(* IEC 61131-3 sources: daoli-st-library/DL_MathData, 454 files *)

(* ---- FC_DL_AccelUnitConvert.st ---- *)
(*==============================================================================
 * 组件名称 (Component)  : FC_DL_AccelUnitConvert
 * 所属子库 (Sublibrary) : DL_MathData ｜ 版本 (Version) : 1.0.0 ｜ 2026-11-23
 * 兼容性   (Platform)   : CODESYS 3.5+ / TwinCAT 3 / 汇川 InoProShop / 施耐德 Machine Expert
 *                         仅依赖 IEC 61131-3 算术运算符，零厂商私有库
 * 功能描述 (Function)   : 加速度单位互转（系数表驱动）：以 m/s² 为中介单位，
 *                         fHub = fValue × kSrc，fResult = fHub ÷ kDst；系数为编译期非零常量，
 *                         纯常量除法，结构性无除零。枚举源/目标越界一律由 CASE ... ELSE
 *                         拦截并返回 0 哨兵（禁静默换算）。
 *                         **重力常数口径**：标准重力加速度 g₀ = 9.80665 m/s²（ISO 80000-3 /
 *                         CGPM 1901 定义值），非本地纬度实测值；本件不做纬度修正。
 * 接口     (Interface)  : 输入 fValue 被换算加速度 [源单位]、eSrc 源单位、eDst 目标单位；
 *                         输出 fConverted 换算结果 [目标单位]、eErrCode（E_DL_AccConvErr）；
 *                         返回值 = 数值可信标志（TRUE = fConverted 可信）。
 * 边界     (Boundary)   : ① 加速度为矢量分量，负值合法（减速 / 反向），不设符号闸。
 *                         ② 单位枚举越域 → 故障级 eInvalidUnit，结果哨兵 0。
 *                         ③ 非有限双判（NaN / ±Inf），命中即故障级 eNonFinite。
 *                         ④ 中介值与结果各复检一次（四段式第四段）。
 *                         ⑤ 零值合法（自由落体失重即 0 g），置信息级 eZeroValue。
 *                         ⑥ 零全局耦合（无 GVL / VAR_EXTERNAL / 物理地址）。
 * 码表     (Codes)      : 本件不占用全局数字码位（R297 零码位范式）；出口为 BOOL + LREAL +
 *                         本文件内 enum E_DL_AccConvErr（全库唯一属主）。
 * 分工声明 (Scope)      : 速度归 FC_DL_SpeedUnitConvert，力归 FC_DL_ForceUnitConvert；
 *                         g 与 m/s² 属加速度量纲，本件专属。
 * 归属     (Ownership)  : E_DL_AccUnit / E_DL_AccConvErr 归属本文件（全库唯一属主，R264）。
 * 红线自检 (Redline)    : R1 ✓ 零 GVL ｜ R2 ✓ 零 %I/%Q ｜ R3 ✓ 纯 IEC ｜ R4 ✓ 非有限双判 +
 *                         CASE ELSE 枚举兜底 + 常量除法无除零 ｜ R5 ✓ 逐行同行双语注释
 *                         R6 ✓ CASE ELSE 兜底（无状态机相位） ｜ R7 N/A（无实例调用）
 * 修订历史 (Revision)   : 2026-11-23  v1.0.0  R78-B2 首版
 * 验收向量 (Acceptance) :
 *   A1 fValue=9.80665, eSrc=eMps2, eDst=eG → 1.0（容差 1E-12）；
 *   A2 fValue=1.0, eSrc=eG, eDst=eMps2 → 9.80665；
 *   A3 fValue=-2.0, eSrc=eMps2, eDst=eG → -0.20394324259558562（负值合法）；
 *   A4 fValue=5.0, eSrc=eMps2, eDst=非法值 7 → 0 哨兵, eInvalidUnit, 返回 FALSE；
 *   A5 fValue=0.0, eSrc=eG, eDst=eMps2 → 0.0, eZeroValue, 返回 TRUE。
 *============================================================================*)

(*-----------------------------------------------------------------------------
 * 枚举: E_DL_AccUnit（加速度单位表，归属本文件，全库唯一属主）
 *----------------------------------------------------------------------------*)
TYPE E_DL_AccUnit :
(
    eMps2 := 0,   // 米每二次方秒（中介单位） / Metre per second squared, hub unit
    eG    := 1    // 标准重力加速度（9.80665 m/s²） / Standard gravity, 9.80665 m/s²
);
END_TYPE

(*-----------------------------------------------------------------------------
 * 枚举: E_DL_AccConvErr（加速度换算出口码；信息级 = 0..9，故障级 = 10 起）
 *----------------------------------------------------------------------------*)
TYPE E_DL_AccConvErr :
(
    eOk          := 0,   // 信息级：换算完成 / Info: conversion completed
    eZeroValue   := 1,   // 信息级：零加速度（失重 / 静止） / Info: zero acceleration, result still trustworthy
    eInvalidUnit := 10,  // 故障级：单位枚举越域 / Fault: unit enum out of domain
    eNonFinite   := 11   // 故障级：输入或结果非有限 / Fault: non-finite input or result
);
END_TYPE

FUNCTION FC_DL_AccelUnitConvert : BOOL
VAR_INPUT
    fValue : LREAL;         // 被换算加速度 [源单位] / Acceleration value in the source unit
    eSrc   : E_DL_AccUnit;  // 源单位枚举 [-] / Source unit enum
    eDst   : E_DL_AccUnit;  // 目标单位枚举 [-] / Destination unit enum
END_VAR
VAR_OUTPUT
    fConverted : LREAL;           // 换算结果 [目标单位] / Converted result in the destination unit
    eErrCode   : E_DL_AccConvErr;  // 出口码 [-] / Outlet code
END_VAR
VAR
    _bBadValue : BOOL;   // 输入非有限标志 [-] / Non-finite input flag
    _fHub      : LREAL;  // 中介加速度值 [m/s²] / Hub acceleration value in metres per second squared
END_VAR
VAR CONSTANT
    DL_ACC_ZERO  : LREAL := 0.0;       // 零基准与零值判定基准 [-] / Zero base
    DL_ACC_MPS2  : LREAL := 1.0;       // m/s² → m/s² 恒等系数 [-] / Hub identity factor
    DL_ACC_G     : LREAL := 9.80665;   // g → m/s² 换算系数（标准重力） / Standard gravity factor
    DL_ACC_EPS   : LREAL := 1.0E-12;   // 零值判定容差 [-] / Zero-detection tolerance
END_VAR

(* —— 段 0：出口预置安全侧 —— *)
FC_DL_AccelUnitConvert := FALSE;                     // 返回值预置不可信 / Return preset not trustworthy
fConverted := DL_ACC_ZERO;                           // 结果哨兵 0 / Result sentinel
eErrCode   := E_DL_AccConvErr.eInvalidUnit;          // 预置最严码 / Preset strictest code

(* —— 段 1：非有限域闸（R79 双判） —— *)
_bBadValue := (fValue <> fValue) OR ((fValue - fValue) <> DL_ACC_ZERO);      // 输入非有限 / Input non-finite
IF _bBadValue THEN
    eErrCode := E_DL_AccConvErr.eNonFinite;          // 故障级码 / Fault-level code
    RETURN;
END_IF

(* —— 段 2：源单位 → 中介 m/s²（CASE ELSE 拦截越域，R6） —— *)
CASE eSrc OF
    E_DL_AccUnit.eMps2 :
        _fHub := fValue * DL_ACC_MPS2;               // 直通 / Hub pass-through
    E_DL_AccUnit.eG :
        _fHub := fValue * DL_ACC_G;                  // g × 9.80665 / Gravity scaled to metres per second squared
ELSE
    _fHub     := DL_ACC_ZERO;                        // 中介值回哨兵 / Hub back to sentinel
    eErrCode  := E_DL_AccConvErr.eInvalidUnit;       // 故障级：源单位越域 / Fault: source unit out of domain
    RETURN;
END_CASE

(* —— 段 3：中介 m/s² → 目标单位（除数为常量，均非零） —— *)
CASE eDst OF
    E_DL_AccUnit.eMps2 :
        fConverted := _fHub / DL_ACC_MPS2;           // ÷1 / Divide by identity
    E_DL_AccUnit.eG :
        fConverted := _fHub / DL_ACC_G;              // ÷9.80665 / Divide by standard gravity factor
ELSE
    fConverted := DL_ACC_ZERO;                       // 结果回哨兵 / Result back to sentinel
    eErrCode   := E_DL_AccConvErr.eInvalidUnit;      // 故障级：目标单位越域 / Fault: destination out of domain
    RETURN;
END_CASE

(* —— 段 4：中介值与结果复检（四段式第四段） —— *)
IF (_fHub <> _fHub) OR ((_fHub - _fHub) <> DL_ACC_ZERO)
    OR (fConverted <> fConverted) OR ((fConverted - fConverted) <> DL_ACC_ZERO) THEN
    fConverted := DL_ACC_ZERO;                       // 复检异常回哨兵 / Recheck failed: sentinel
    eErrCode   := E_DL_AccConvErr.eNonFinite;        // 故障级码 / Fault-level code
    RETURN;
END_IF

(* —— 段 5：成功出口（零值单列信息码） —— *)
IF (fValue < DL_ACC_EPS) AND (fValue > -DL_ACC_EPS) THEN
    eErrCode := E_DL_AccConvErr.eZeroValue;          // 信息级：零加速度 / Info: zero acceleration
ELSE
    eErrCode := E_DL_AccConvErr.eOk;                 // 信息级：换算完成 / Info: conversion completed
END_IF
FC_DL_AccelUnitConvert := TRUE;                      // 换算有效 / Conversion valid
END_FUNCTION

(* ---- FC_DL_AngleUnitConvert.st ---- *)
// ==============================================================================
// 组件名 Component  : FC_DL_AngleUnitConvert
// 分类   Category   : DL_MathData
// 前缀   Naming     : FC_DL_ ｜ b/f/e 类型前缀制（R265）
// 版本   Version    : 1.0.0
// 复杂度 Complexity  : 低
// 功能   Purpose    : 角度单位换算（度 / 弧度 / 梯度）：统一转 rad 中间量
//                      再转目标单位，任意两单位直换（deg → grad 系数
//                      200/180 经 rad 中转自动成立）。非有限输入拒绝
//                      （bValid = FALSE、fOut = 0.0）。
// 开源溯源 Origin    : 道莅原创（角度单位定义为公开计量常识，本实现
//                      clean-room，未复制任何源码行；与 TempUnitConvert /
//                      PressUnitConvert / FlowUnitConvert 同族单位换算
//                      组织口径）
// 许可证 License    : MIT
// 参考   Reference  : IEC 61131-3:2013 §6.6.2 CASE 语义；角度单位换算公开
//                      计量定义（借定义，不抄实现）
// 平台   Platform   : 纯 IEC 61131-3（CASE / LREAL 四则），三平台通用
// 依赖   Depends    : 无（零委托、零库件；换算系数常量预乘，运行期零除法）
// 分工声明 Split     : FC_DL_AngleDiffWrap（角差归一）与 FC_DL_WrapAngleDeg
//                      （角度回绕）与本件互引；本件只做单位换算（不改
//                      角度主值、不回绕），归一 / 回绕语义归各自属主（R216）。
// 归属 Ownership     : E_DL_AngUnit 属主为本文件（全库唯一定义，R264）；
//                      引用件只引用不重声明。
// ------------------------------------------------------------------
// 边界 Boundary     :
//   一 非有限闸：fVal 为 NaN（自反判 x <> x）或 ±Inf（差值自反判
//      (x - x) <> (x - x)）或幅值越 1e30 上界 → bValid = FALSE、
//      fOut = 0.0 早退（故障级 0749，R272 非有限防护）；
//   二 零除法面：四向系数全部预乘为常量（PI/180、180/PI、PI/200、
//      200/PI 编译期落定），运行期无除法（除零面结构性消除）；
//   三 枚举闸：eFrom / eTo 非法枚举值（CASE ELSE 兜底）→ bValid =
//      FALSE、fOut = 0.0 早退（与 0749 同形出口合并一码，R90 反证句：
//      现有输出组合不可区分两场景）；
//   四 纯函数：无记忆量、无定时器、无边沿实例，每调用重算；
//   五 无全局、无外部变量、无物理地址。
// 错误码 Codes      :
//   16#0001_0749【故障级】输入非有限或枚举非法（bValid = FALSE、
//                fOut = 0.0 早退）
//   注：本件引脚契约按任务定稿无独立 eErr 出口，故障语义经
//   bValid = FALSE + fOut = 0.0 组合表达。
// 验收 Acceptance   :
//   算法已证（脚本）：未跑 ｜ 编译器已证（三平台）：未跑
//   V1 180 deg → rad = 3.14159265358979；V2 1 rad → deg = 57.2957795
//   V3 200 grad → rad = 3.14159265358979；V4 180 deg → grad = 200（200/180 系数）
//   V5 fVal = NaN → bValid = FALSE、fOut = 0.0
//   V6 eFrom 非法枚举 → bValid = FALSE、fOut = 0.0
// 修订记录 Revision  :
//   2026-11-22  v1.0.0  R65 首版（批 2 · 序号 7）
// ==============================================================================
TYPE E_DL_AngUnit :
(
    eDeg  := 0, // 度 [deg]，一周 360 / degrees, 360 per turn
    eRad  := 1, // 弧度 [rad]，一周 2*PI / radians, two pi per turn
    eGrad := 2  // 梯度 [grad]，一周 400 / gradians, 400 per turn
);
END_TYPE

FUNCTION FC_DL_AngleUnitConvert : BOOL
VAR_INPUT
    fVal  : LREAL;               // 输入角值 [源单位] / the input angle in the source unit
    eFrom : E_DL_AngUnit;        // 源单位枚举 [单位] / the source unit
    eTo   : E_DL_AngUnit;        // 目标单位枚举 [单位] / the target unit
END_VAR
VAR_OUTPUT
    fOut   : LREAL;              // 输出角值 [目标单位]，无效时 0.0 / the output angle in the target unit, zero when invalid
    bValid : BOOL;               // 结果可用 [-]，非有限或枚举非法为 FALSE / the validity flag
END_VAR
VAR
    fRad : LREAL;                // 中间弧度量 [rad]（统一中转）/ the intermediate radian value
END_VAR
VAR CONSTANT
    DL_AUC_D2R  : LREAL := 0.0174532925199433;   // 度 → 弧度系数 [rad/deg]，PI/180 预乘 / the deg to rad factor, pi over one eighty
    DL_AUC_R2D  : LREAL := 57.2957795130823;     // 弧度 → 度系数 [deg/rad]，180/PI 预乘 / the rad to deg factor
    DL_AUC_G2R  : LREAL := 0.0157079632679490;   // 梯度 → 弧度系数 [rad/grad]，PI/200 预乘 / the grad to rad factor, pi over two hundred
    DL_AUC_R2G  : LREAL := 63.6619772367581;     // 弧度 → 梯度系数 [grad/rad]，200/PI 预乘 / the rad to grad factor
    DL_AUC_FMAX : LREAL := 1.0E30;               // 非有限筛查幅值上限 [源单位] / the finiteness screening cap
END_VAR

// 段 1｜返回值与全部出口预置（R45 四段式第一段）/ segment 1, the preset of the return and all outlets
FC_DL_AngleUnitConvert := FALSE; // 返回值预置假 / preset the return false
fOut   := 0.0;                   // 输出预置零 [目标单位] / preset the output zero
bValid := FALSE;                 // 有效标志预置假 / preset the validity false
fRad   := 0.0;                   // 中间量预置零 [rad] / preset the intermediate zero

// 段 2｜非有限闸（边界一：NaN 自反判 + Inf 差值自反判 + 幅值上界，R272）/ segment 2, the non finite gate
IF (fVal <> fVal) OR ((fVal - fVal) <> 0.0) OR (ABS(fVal) > DL_AUC_FMAX) THEN // 输入非有限 / the input non finite
    fOut   := 0.0;               // 输出归零 [目标单位] / zero the output
    bValid := FALSE;             // 故障级 0749：拒绝换算 / refuse the conversion
    RETURN;                      // 早退 / early return
END_IF

// 段 3｜源单位归一到 rad（边界三：CASE 带 ELSE 兜底）/ segment 3, the source unit normalization to radians
CASE eFrom OF
    E_DL_AngUnit.eDeg:           // 度 → rad / degrees to radians
        fRad := fVal * DL_AUC_D2R; // 乘 PI/180 系数 [rad] / multiply the deg to rad factor
    E_DL_AngUnit.eRad:           // 弧度直通 / radians pass through
        fRad := fVal;            // 中转量即输入 [rad] / the intermediate is the input
    E_DL_AngUnit.eGrad:          // 梯度 → rad / gradians to radians
        fRad := fVal * DL_AUC_G2R; // 乘 PI/200 系数 [rad] / multiply the grad to rad factor
    ELSE                         // 非法枚举拦截（边界三）/ an illegal enumeration
        fOut   := 0.0;           // 输出归零 / zero the output
        bValid := FALSE;         // 故障级 0749 同形出口（R90 合并）/ the merged fault outlet
        RETURN;                  // 早退 / early return
END_CASE

// 段 4｜rad 转目标单位（边界三：CASE 带 ELSE 兜底）/ segment 4, the radians to the target unit
CASE eTo OF
    E_DL_AngUnit.eDeg:           // rad → 度 / radians to degrees
        fOut := fRad * DL_AUC_R2D; // 乘 180/PI 系数 [deg] / multiply the rad to deg factor
    E_DL_AngUnit.eRad:           // rad 直通 / radians pass through
        fOut := fRad;            // 输出即中转量 [rad] / the output is the intermediate
    E_DL_AngUnit.eGrad:          // rad → 梯度 / radians to gradians
        fOut := fRad * DL_AUC_R2G; // 乘 200/PI 系数（deg → grad 经此链自动得 200/180）[grad] / the rad to grad factor
    ELSE                         // 非法枚举拦截（边界三）/ an illegal enumeration
        fOut   := 0.0;           // 输出归零 / zero the output
        bValid := FALSE;         // 故障级 0749 同形出口（R90 合并）/ the merged fault outlet
        RETURN;                  // 早退 / early return
END_CASE

// 段 5｜统一出口 / segment 5, the unified outlet
bValid := TRUE;                  // 结果可用 / the result usable
FC_DL_AngleUnitConvert := TRUE;  // 返回成功 / return success
END_FUNCTION

(* ---- FC_DL_AreaUnitConvert.st ---- *)
(*==============================================================================
 * 组件名称 (Component)  : FC_DL_AreaUnitConvert
 * 所属子库 (Sublibrary) : DL_MathData
 * 当前版本 (Version)    : 1.0.0
 * 兼容性   (Platform)   : CODESYS 3.5+ / TwinCAT 3 / 汇川 InoProShop / 施耐德 Machine Expert
 *                         仅依赖 IEC 61131-3 算术运算符，零厂商私有库
 * 功能描述 (Function)   : 面积单位换算（系数表驱动）：以平方米（m²）为中介单位，
 *                         fHub = fValue × kSrc，fResult = fHub ÷ kDst；系数为编译期
 *                         非零常量，纯常量除法，结构性无除零。
 *                         **量纲警告**：面积系数是长度系数的平方（mm² = 1E-6 m²、
 *                         ft² = 0.09290304 m²），不可与长度系数混用；本件显式使用
 *                         平方后的常量，禁止由长度族推导。
 *                         面积非负：负值判故障级 eNegativeValue 并回哨兵 0。
 * 接口     (Interface)  : 输入 fValue 被换算面积 [源单位]、eSrc 源单位、eDst 目标单位；
 *                         输出 fConverted 换算结果 [目标单位]、eErrCode（E_DL_AreaConvErr）；
 *                         返回值 = bValid 数值可信标志（TRUE = fConverted 可信）。
 * 边界     (Boundary)   : ① 属主边界：只做单位换算，不做体积 = 面积 × 行程 的推导。
 *                         ② 单位枚举越域 → 故障级 eInvalidUnit，结果哨兵 0。
 *                         ③ 非有限双判，命中即故障级 eNonFinite。
 *                         ④ 负面积 → 故障级 eNegativeValue（拒绝，不钳位）。
 *                         ⑤ 零值合法（info 级 eZeroValue）。结果与中介值各复检一次。
 *                         ⑥ 极小量纲提示：mm² 值域可极大（1 m² = 1E6 mm²），LREAL 尾数
 *                         53 位，最大可表 1.8E308，无溢出风险；但仍做非有限复检。
 *                         ⑦ 零全局耦合（无 GVL / VAR_EXTERNAL / 物理地址）。
 * 分工声明 (Scope)      : 与 `FC_DL_LengthUnitConvert` 分工：长度归那件，本件自带平方系数，
 *                         严禁调用长度件再平方（会引入两次舍入误差并破坏枚举域闸）。
 * 来源标签 (Source Tag) : 开源溯源：lgf-math 换算系数（公开物理常数，clean-room 重写）；许可证 MIT（仅参考语义，代码原创）
 * 码表     (Codes)      : 本件不占用全局数字码位；出口为 BOOL + LREAL +
 *                         本文件内定义 enum E_DL_AreaConvErr（全库唯一）。
 * 红线自检 (Redline)    : R1 ✓ 零 GVL/VAR_EXTERNAL ｜ R2 ✓ 零 %I/%Q/%M ｜ R3 ✓ 纯 IEC 61131-3
 *                         R4 ✓ 非有限双判 + 枚举域闸 + 常量除法无除零 + 负值拒绝 ｜ R5 ✓ 声明逐行同行双语注释
 *                         R6 N/A（纯函数无状态机） ｜ R7 N/A（无实例调用）
 * 修订历史 (Revision)   : 2026-11-23  v1.0.0  R77 首版（批次 B2 · 序号 14）
 * 验收向量 (Acceptance) : ① fValue=1.0, eSrc=eM2, eDst=eMm2 → 1×1.0 = 1 m2,
 *                         ÷1E-6 = 1000000.0 mm2（容差 1E-3）；
 *                         ② fValue=1.0, eSrc=eFt2, eDst=eM2 → 1×0.09290304 = 0.09290304 m2；
 *                         ③ fValue=1000000.0, eSrc=eMm2, eDst=eM2 → 1000000×1E-6 = 1.0 m2；
 *                         ④ fValue=-1.0, eSrc=eM2, eDst=eFt2 → 返回 FALSE, 0, eNegativeValue。
 *==============================================================================*)

(*-----------------------------------------------------------------------------
 * 枚举: E_DL_AreaUnit（面积单位表，归属 DL_MathData，与本件同文件，全库唯一属主）
 *----------------------------------------------------------------------------*)
TYPE E_DL_AreaUnit :
(
    eMm2 := 0,   // 平方毫米（1E-6 m2） / Square millimetre
    eM2  := 1,   // 平方米（中介单位） / Square metre, hub unit
    eFt2 := 2    // 平方英尺（0.09290304 m2，= 0.3048^2） / Square foot
);
END_TYPE

(*-----------------------------------------------------------------------------
 * 枚举: E_DL_AreaConvErr（面积换算错误码）
 *----------------------------------------------------------------------------*)
TYPE E_DL_AreaConvErr :
(
    eOk            := 0,   // 信息级：换算完成 / Info: conversion completed
    eZeroValue     := 1,   // 信息级：输入为零（合法） / Info: zero input, legal
    eInvalidUnit   := 2,   // 故障级：单位枚举越域 / Fault: unit enum out of domain
    eNonFinite     := 3,   // 故障级：输入非有限 / Fault: non-finite input
    eNegativeValue := 4    // 故障级：负面积 / Fault: negative area
);
END_TYPE

FUNCTION FC_DL_AreaUnitConvert : BOOL
VAR_INPUT
    fValue : LREAL;          // 被换算面积值 [源单位] / Area value in source unit
    eSrc   : E_DL_AreaUnit;  // 源单位枚举 [-] / Source unit enum
    eDst   : E_DL_AreaUnit;  // 目标单位枚举 [-] / Destination unit enum
END_VAR
VAR_OUTPUT
    fConverted : LREAL;            // 换算结果 [目标单位] / Converted result
    eErrCode   : E_DL_AreaConvErr; // 错误码出口 [-] / Error code outlet
END_VAR
VAR
    _bNonFin : BOOL;   // 输入非有限当拍标志 [-] / Non-finite input flag
    _fHub    : LREAL;  // 中介面积值 [m2] / Hub area value in square metres
END_VAR
VAR CONSTANT
    DL_AUC_MM2  : LREAL := 1.0E-6;      // mm2 → m2 换算系数（0.001^2） [m2/mm2] / square millimetre to square metre factor
    DL_AUC_M2   : LREAL := 1.0;         // m2 → m2 恒等系数 [m2/m2] / square metre identity factor
    DL_AUC_FT2  : LREAL := 0.09290304;  // ft2 → m2 换算系数（0.3048^2） [m2/ft2] / square foot to square metre factor
    DL_AUC_ZERO : LREAL := 0.0;         // 零值与非有限判零基准 [-] / Zero and non-finite base
END_VAR

(* —— 段 0：出口预置安全值 —— *)
FC_DL_AreaUnitConvert := FALSE;                    // 返回值预置无效 / Return preset invalid
fConverted := DL_AUC_ZERO;                         // 结果哨兵 0 / Result sentinel
eErrCode   := E_DL_AreaConvErr.eInvalidUnit;       // 预置最严码 / Preset strictest code

(* —— 段 1：非有限域闸（R79 双判） —— *)
_bNonFin := (fValue <> fValue) OR ((fValue - fValue) <> DL_AUC_ZERO);   // 非有限判定 / Non-finite test
IF _bNonFin THEN
    eErrCode := E_DL_AreaConvErr.eNonFinite;       // 故障级码 / Fault-level code
    RETURN;
END_IF

(* —— 段 2：负面积域闸 —— *)
IF fValue < DL_AUC_ZERO THEN
    eErrCode := E_DL_AreaConvErr.eNegativeValue;   // 故障级码 / Fault-level code
    RETURN;
END_IF

(* —— 段 3：源单位 → 中介平方米 —— *)
IF eSrc = E_DL_AreaUnit.eMm2 THEN
    _fHub := fValue * DL_AUC_MM2;                  // mm2 × 1E-6 / square millimetre scaled
ELSIF eSrc = E_DL_AreaUnit.eM2 THEN
    _fHub := fValue * DL_AUC_M2;                   // m2 直通 / square metre pass-through
ELSIF eSrc = E_DL_AreaUnit.eFt2 THEN
    _fHub := fValue * DL_AUC_FT2;                  // ft2 × 0.09290304 / square foot scaled
ELSE
    RETURN;                                        // 源单位越域 / Source unit out of domain
END_IF

(* —— 段 4：中介平方米 → 目标单位（常量除法，分母非零） —— *)
IF eDst = E_DL_AreaUnit.eMm2 THEN
    fConverted := _fHub / DL_AUC_MM2;              // ÷1E-6（放大 1e6，注意量纲） / Divide by square millimetre factor
ELSIF eDst = E_DL_AreaUnit.eM2 THEN
    fConverted := _fHub / DL_AUC_M2;               // ÷1 / Divide by identity
ELSIF eDst = E_DL_AreaUnit.eFt2 THEN
    fConverted := _fHub / DL_AUC_FT2;              // ÷0.09290304 / Divide by square foot factor
ELSE
    eErrCode   := E_DL_AreaConvErr.eInvalidUnit;   // 目标单位越域 / Destination out of domain
    fConverted := DL_AUC_ZERO;
    RETURN;
END_IF

(* —— 段 5：结果非有限复检兜底（量级放大 1e6 后必须复检） —— *)
IF (fConverted <> fConverted) OR ((fConverted - fConverted) <> DL_AUC_ZERO) THEN
    fConverted := DL_AUC_ZERO;                     // 复检异常回哨兵 / Recheck failed: sentinel
    eErrCode   := E_DL_AreaConvErr.eNonFinite;     // 故障级码 / Fault-level code
    RETURN;
END_IF

(* —— 段 6：成功出口 —— *)
IF fValue = DL_AUC_ZERO THEN
    eErrCode := E_DL_AreaConvErr.eZeroValue;       // 信息级：零值 / Info: zero value
ELSE
    eErrCode := E_DL_AreaConvErr.eOk;              // 信息级成功 / Info success
END_IF
FC_DL_AreaUnitConvert := TRUE;                     // 换算有效 / Conversion valid

END_FUNCTION

(* ---- FC_DL_CharCodeConvert.st ---- *)
(*
    FC_DL_CharCodeConvert —— 单字符 ↔ 字符码双向换算原子
    ------------------------------------------------------------------
    组件名称  : FC_DL_CharCodeConvert
    分类      : DL_MathData / CharCode
    前缀      : FC_DL_
    版本      : 1.0.0
    溯源      : IEC 61131-3 标准语义的道莅防御性实现（单字符与码值的
                双向映射原子，映射内核 = 定长字符表 + 标准 MID / FIND
                检索，零内建转换链依赖）；实现 / 引脚名 / 码位 100% 自有；
                clean-room 声明 —— 零代码行复制，无闭源参考。
    平台      : 纯 IEC 61131-3（Standard.library: LEN / MID / FIND），
                CODESYS 3.5 / TwinCAT 3 / InoProShop / Machine Expert 通用
    作者      : 道莅代码库 · PLC编程专家（R72 构建轮 · 批 2 · 序号 4）
    ------------------------------------------------------------------
    功能说明  : 单字符与字符码（0~255）双向换算。真实工况：HMI 键盘映射、
                协议字符组装、标签打印机字符转义。选向由 eMode 枚举显式
                给出，未选方向出口置确定值（空串 / 0），绝不残留旧值。
                判据链顺序：
                ① eCharToCode 向：串长域闸（LEN <> 1 → 拒收信息级，空串 /
                   多字符同样拒收）→ LO / HI 双表 FIND 检索（先 LO 后 HI，
                   命中即回码值）→ 双表全未命中 → 防御性拒收（结构性不可达，
                   表覆盖 1..255 全字节）；
                ② eCodeToChar 向：码域闸（uCodeIn > 255 → 故障级早退）→
                   码 0 = 串终结符，回执空串（忠实语义，声明口径）→ 码
                   1..127 查 LO 表（位置 = 码值）、码 128..255 查 HI 表
                   （位置 = 码值 − 127）；
                ③ 选向枚举漏项由 CASE ELSE 兜底（拒收信息级，双出口置
                   确定值）。
                扩展 ASCII 披露（128~255）：本件只保证**码值回执**的字节级
                正确性，不保证三平台对 $80~$FF 的渲染 / 显示一致（字体与
                代码页差异属显示层语义），头注释声明披露。
                交付门槛（R64 口径）：MID / FIND 对 $80~$FF 字节的检索行为
                须在 CODESYS / TwinCAT / InoProShop 三平台各编译验证一次。
    错误码    : 16#0002_3906 码域越界（uCodeIn > 255），双出口置确定值空串/0
                            —— 故障级
                16#0002_3907 串长域闸拒收（LEN <> 1，空串 / 多字符同拒）
                            —— 信息级，不置 bError（R45）
                16#0002_3908 选向枚举漏项（CASE ELSE 兜底拒收）—— 信息级，
                            不置 bError
                加码反证句（R90）：3906 由「故障级 + 双出口确定值」唯一观测；
                3907 与 3908 在输出组合上不可分（同为拒收），但成因互斥
                （串长 vs 选向）且调用方可自证入参，故按成因分立两码，
                拒绝合并导致选向错误被误报为串长错误。
    码位总账  : 16#0002_3906 用 ｜ 16#0002_3907 用 ｜ 16#0002_3908 用
    状态机    : 无顺序状态机；选向用 CASE + ELSE 兜底（非法枚举值拦截），
                枚举成员初值一律 :=（红线 4）
    边界与披露: 一 无定时器 / 无沿检测实例 / 无数组下标 / 无除法，周期安全
                   规则 N/A；
                二 零全局变量、零 VAR_EXTERNAL、零物理地址；
                三 域闸逐项点名（R272）：uCodeIn 码域闸覆盖 0~255 全段
                   （0 与 255 两端点各推一条向量）；sCharIn 串长闸覆盖
                   0 / 1 / 多字符三态；
                四 双出口默认值纪律：未选向 / 拒收路径 sCharOut = ''、
                   uCodeOut = 0 确定值，绝不残留旧值（R256）；
                五 字符表覆盖声明：LO 表覆盖码 1..127、HI 表覆盖码 128..255、
                   码 0 按串终结符语义回执空串——三段并起覆盖 0..255 全域，
                   无缺口；
                六 与 FC_DL_HexStringToBytes / FC_DL_DwordToHexString 分工
                   互引：那两件是文本 ↔ 字节块，本件是单字符 ↔ 码值原子，
                   不互代；
                七 依赖声明：仅 Standard.library（LEN / MID / FIND），
                   零厂商方言。
    验收向量  : V1 eCodeToChar，uCodeIn = 0 → 空串（终结符语义）；
                V2 eCodeToChar，uCodeIn = 65 → 'A'；V3 eCodeToChar，
                uCodeIn = 255 → '$FF' 字符；V4 eCodeToChar，uCodeIn = 256
                → 3906 故障级；V5 eCharToCode，'A' → 65；
                V6 eCharToCode，'' 或 'AB' → 3907 拒收；
                V7 eCharToCode，' '（空格，码 32）→ 32。
                算法已证（脚本）：未跑 ｜ 编译器已证（三平台）：未跑
    修订记录  : 2026-11-23 v1.0.0 首次入库（R72 构建轮 · 批 2 · 序号 4）
*)
TYPE E_DL_CharCodeMode :
(
    eCharToCode := 0,                      // 选向：字符 → 码值 / the direction char to code
    eCodeToChar := 1                       // 选向：码值 → 字符 / the direction code to char
);
END_TYPE

FUNCTION FC_DL_CharCodeConvert : BOOL
VAR_INPUT
    eMode    : E_DL_CharCodeMode;          (* 换算方向选向，[选向枚举] / the conversion direction selector *)
    sCharIn  : STRING;                     (* 字符输入（eCharToCode 向用），[串]，串长闸限 1 字符 / the char input, gated to one char *)
    uCodeIn  : UINT;                       (* 码值输入（eCodeToChar 向用），[码]，域 0~255 / the code input, domain 0 to 255 *)
END_VAR
VAR_OUTPUT
    sCharOut  : STRING(1);                 (* 字符出口（未选向 / 拒收时为空串确定值）[串] / the char outlet, empty when rejected *)
    uCodeOut  : UINT;                      (* 码值出口（未选向 / 拒收时为 0 确定值）[码] / the code outlet, zero when rejected *)
    bValid    : BOOL;                      (* 输出可用标志，拒收 / 故障为 FALSE / the outputs usable flag *)
    bError    : BOOL;                      (* 故障标志，仅故障级码置位（R45 配对）/ the fault flag *)
    nInfoCode : UDINT;                     (* 信息 / 错误码，0 = 正常 / the info or error id *)
END_VAR
VAR CONSTANT
    DL_CHC_TAB_LO : STRING(127) := '$01$02$03$04$05$06$07$08$09$0A$0B$0C$0D$0E$0F$10$11$12$13$14$15$16$17$18$19$1A$1B$1C$1D$1E$1F !"$24%&$27()*+,-./0123456789:;<=>?@ABCDEFGHIJKLMNOPQRSTUVWXYZ[\]^_`abcdefghijklmnopqrstuvwxyz{|}~$7F'; (* 码 1..127 字符表（位置 p = 码 p），$24 = '$'，$27 = ''' / the low char table, position p equals code p *)
    DL_CHC_TAB_HI : STRING(128) := '$80$81$82$83$84$85$86$87$88$89$8A$8B$8C$8D$8E$8F$90$91$92$93$94$95$96$97$98$99$9A$9B$9C$9D$9E$9F$A0$A1$A2$A3$A4$A5$A6$A7$A8$A9$AA$AB$AC$AD$AE$AF$B0$B1$B2$B3$B4$B5$B6$B7$B8$B9$BA$BB$BC$BD$BE$BF$C0$C1$C2$C3$C4$C5$C6$C7$C8$C9$CA$CB$CC$CD$CE$CF$D0$D1$D2$D3$D4$D5$D6$D7$D8$D9$DA$DB$DC$DD$DE$DF$E0$E1$E2$E3$E4$E5$E6$E7$E8$E9$EA$EB$EC$ED$EE$EF$F0$F1$F2$F3$F4$F5$F6$F7$F8$F9$FA$FB$FC$FD$FE$FF'; (* 码 128..255 字符表（位置 p = 码 127 + p），只保证码值回执不保证显示 / the high char table, position p equals code 127 plus p *)
    DL_CHC_ONE    : INT  := 1;             (* 检索步进与串长基准 [个] / the search step and the length base *)
    DL_CHC_SPLIT  : UINT := 127;           (* LO / HI 表码值分界 [码] / the code split between the tables *)
    DL_CHC_CMAX   : UINT := 255;           (* 码域上界 [码] / the code domain upper bound *)
    DL_CHC_ZERO   : UINT := 0;             (* 码零哨兵（终结符语义）[码] / the zero code sentinel *)
    DL_CHC_ZEROI  : INT  := 0;             (* 检索未命中哨兵 [位置] / the not found sentinel *)
END_VAR
VAR
    nLen  : INT;                           (* 输入串长 [个] / the input string length *)
    nPos  : INT;                           (* FIND 检索命中位置（LO 表）[位置] / the FIND hit position in the low table *)
    nPosH : INT;                           (* FIND 检索命中位置（HI 表）[位置] / the FIND hit position in the high table *)
END_VAR

// 段 1｜返回值与双出口预置（统一出口预置，R256）/ segment 1, preset the return and the dual outlets
FC_DL_CharCodeConvert := FALSE;          // 故障缺省返回不可用 / the fault default is unusable
sCharOut  := '';                         // 字符出口预置空串确定值 / preset the char outlet to the empty string
uCodeOut  := DL_CHC_ZERO;                // 码值出口预置零确定值 / preset the code outlet to zero
bValid    := FALSE;                      // 可用标志预清零 / preset the usable flag false
bError    := FALSE;                      // 故障标志预清零 / preset the fault flag false
nInfoCode := 0;                          // 码位预置无错 / preset the code to zero
nLen  := 0;                              // 串长中间量清零 / clear the length temporary
nPos  := DL_CHC_ZEROI;                   // 检索位置清零 / clear the hit position
nPosH := DL_CHC_ZEROI;                   // 检索位置清零 / clear the hit position

// 段 2｜选向分发（CASE + ELSE 兜底，非法枚举值拦截，红线 4）/ segment 2, the direction dispatch with the ELSE guard
CASE eMode OF

    E_DL_CharCodeMode.eCharToCode:       // 字符 → 码值向 / the char to code direction
        nLen := LEN(sCharIn);            // 串长闸取样 / sample the input length
        IF nLen <> DL_CHC_ONE THEN       // 空串或多字符一律拒收（串长域闸）/ empty or multi char rejected
            nInfoCode := 16#0002_3907;   // 信息级：串长闸拒收 / info level: the length gate rejection
            bError := FALSE;             // 信息级不置故障（R45）/ info level never raises a fault
            bValid := FALSE;             // 输出不可用 / the outputs unusable
            sCharOut := '';              // 双出口确定值（R256）/ the deterministic outlets
            uCodeOut := DL_CHC_ZERO;     // 双出口确定值 / the deterministic outlets
            RETURN;                      // 结构早退 / structural exit
        END_IF
        nPos := FIND(DL_CHC_TAB_LO, sCharIn); // LO 表检索（位置 p = 码 p）/ search the low table
        IF nPos > DL_CHC_ZEROI THEN      // LO 表命中 / a low table hit
            uCodeOut := INT_TO_UINT(nPos); // 码值 = 位置 / the code equals the position
        ELSE                             // LO 未命中转 HI 表 / fall through to the high table
            nPosH := FIND(DL_CHC_TAB_HI, sCharIn); // HI 表检索（位置 p = 码 127 + p）/ search the high table
            IF nPosH > DL_CHC_ZEROI THEN // HI 表命中 / a high table hit
                uCodeOut := INT_TO_UINT(nPosH + UINT_TO_INT(DL_CHC_SPLIT)); // 码值 = 位置 + 127 / the code equals position plus 127
            ELSE                         // 双表全未命中（表覆盖 1..255 全字节，结构性不可达防御收口）/ both tables missed, unreachable
                nInfoCode := 16#0002_3907; // 信息级：检索失败按拒收口径 / info level: the search failure rejection
                bValid := FALSE;         // 输出不可用 / unusable
                sCharOut := '';          // 双出口确定值 / the deterministic outlets
                uCodeOut := DL_CHC_ZERO; // 双出口确定值 / the deterministic outlets
                RETURN;                  // 结构早退 / exit
            END_IF
        END_IF
        bValid := TRUE;                  // 换算成功 / the conversion succeeded

    E_DL_CharCodeMode.eCodeToChar:       // 码值 → 字符向 / the code to char direction
        IF uCodeIn > DL_CHC_CMAX THEN    // 码域闸（>255 越域）/ the code domain gate
            nInfoCode := 16#0002_3906;   // 故障级：码域越界 / fault level: the code domain violation
            bError := TRUE;              // R45 配对置故障标志 / paired with the fault flag
            bValid := FALSE;             // 输出不可用 / unusable
            sCharOut := '';              // 双出口确定值 / the deterministic outlets
            uCodeOut := DL_CHC_ZERO;     // 双出口确定值 / the deterministic outlets
            RETURN;                      // 结构早退 / exit
        END_IF
        uCodeOut := uCodeIn;             // 码值回执（选向确认）/ echo the code
        IF uCodeIn = DL_CHC_ZERO THEN    // 码 0 = 串终结符，忠实回执空串 / code zero is the terminator, faithful empty
            sCharOut := '';              // 空串出口 / the empty outlet
        ELSIF uCodeIn <= DL_CHC_SPLIT THEN // 码 1..127 查 LO 表 / the low table range
            nPos := UINT_TO_INT(uCodeIn); // 位置 = 码值（LO 表 1 起）/ the position equals the code
            sCharOut := MID(DL_CHC_TAB_LO, nPos, DL_CHC_ONE); // 取单字符 / pick the single char
        ELSE                             // 码 128..255 查 HI 表 / the high table range
            nPos := UINT_TO_INT(uCodeIn) - UINT_TO_INT(DL_CHC_SPLIT); // 位置 = 码值 − 127 / the position equals code minus 127
            sCharOut := MID(DL_CHC_TAB_HI, nPos, DL_CHC_ONE); // 取单字符 / pick the single char
        END_IF
        bValid := TRUE;                  // 换算成功 / the conversion succeeded

    ELSE                                 // 选向枚举漏项兜底（红线 4）/ the unknown direction guard
        nInfoCode := 16#0002_3908;       // 信息级：选向未知拒收 / info level: the unknown direction rejection
        bError := FALSE;                 // 信息级不置故障（R45）/ info level never raises a fault
        bValid := FALSE;                 // 输出不可用 / unusable
        sCharOut := '';                  // 双出口确定值 / the deterministic outlets
        uCodeOut := DL_CHC_ZERO;         // 双出口确定值 / the deterministic outlets

END_CASE

// 段 3｜统一出口 / segment 3, the unified outlet
FC_DL_CharCodeConvert := bValid;         // 返回值与 bValid 同源（R191 名实双出口）/ the return shares its source with bValid
END_FUNCTION

(* ---- FC_DL_CircleFit3Pt.st ---- *)
(*==============================================================================
 * 组件名称 (Component)  : FC_DL_CircleFit3Pt
 * 所属子库 (Sublibrary) : DL_MathData
 * 当前版本 (Version)    : 1.0.0
 * 兼容性   (Platform)   : CODESYS 3.5+ / TwinCAT 3 / 汇川 InoProShop / 施耐德 Machine Expert
 *                         仅依赖 Standard.library（SQRT / ABS），零厂商私有库
 * 功能描述 (Function)   : 三点定圆（外接圆解析解，代数行列式法）：
 *                           D  = 2×[x1(y2−y3) + x2(y3−y1) + x3(y1−y2)]
 *                           Ux = [(x1²+y1²)(y2−y3) + (x2²+y2²)(y3−y1)
 *                                 + (x3²+y3²)(y1−y2)] ÷ D
 *                           Uy = [(x1²+y1²)(x3−x2) + (x2²+y2²)(x1−x3)
 *                                 + (x3²+y3²)(x2−x1)] ÷ D
 *                           R  = SQRT((x1−Ux)² + (y1−Uy)²)
 *                         |D| < 共线容差判三点共线（叉积绝对值判据），拒绝并置
 *                         故障码 eCollinear（防除零前置闸，规格指定）；非有限
 *                         输入 → 故障码 eNonFinite，输出哨兵 0。
 * 接口     (Interface)  : 输入 fX1/fY1/fX2/fY2/fX3/fY3 三点坐标 [mm]；
 *                         输出 fCx 圆心横坐标 [mm]、fCy 圆心纵坐标 [mm]、
 *                         fR 半径 [mm]、eErrCode 错误码（E_DL_CircFitErr）、
 *                         返回值 = 拟合有效标志（BOOL）。
 * 边界     (Boundary)   : ① **属主边界（写死）：本件只做三点定圆解析解，不做
 *                         多点最小二乘拟合、不做圆度评价**；多点拟合归
 *                         统计类件。
 *                         ② 共线闸：|D| = |2×叉积| < DL_CFT_COLMIN → 拒算
 *                         （D 作除数前置判，结构性无除零）；容差量纲随坐标
 *                         单位（mm 口径下 1E-9 对应亚纳米叉积面积），头注释
 *                         声明为「近共线拒算域」，非严格共线唯一判据。
 *                         ③ 非有限判据（R79 双判）：六坐标逐一 NaN 自反
 *                         x <> x 与 Inf 差自减 (x−x) <> (x−x)。
 *                         ④ R 非负结构性保证：平方和开方，无负数开方路径。
 *                         ⑤ 输出预置哨兵 0 早退（四段式：预置→域闸→内核→
 *                         结果复检），任何早退路径前输出已确定。
 *                         ⑥ 零全局耦合（无 GVL / VAR_EXTERNAL / 物理地址）。
 * 分工声明 (Scope)      : 与 `FC_DL_CalcDistance3D` 分工：距离原语归那件、
 *                         三点定圆归本件；本件 SQRT 只用于半径合成（属主
 *                         内核例外申报：本件为圆拟合内核属主）。
 * 来源标签 (Source Tag) : 自研线（外接圆行列式公式为公开解析几何定义 clean-room）
 * 码表     (Codes)      : 本件不占用任何全局数字码位。出口为 BOOL 返回 +
 *                         LREAL 三值 + ENUM 错误码；数字码位待主控收口阶段
 *                         统一派号。
 * 红线自检 (Redline)    : R1 ✓ 零 GVL/VAR_EXTERNAL ｜ R2 ✓ 零 %I/%Q/%M ｜ R3 ✓ 纯 IEC 61131-3
 *                         R4 ✓ 共线前置闸防除零 + 非有限双判 + 哨兵早退 ｜ R5 ✓ 声明逐行同行双语注释
 *                         R6 N/A（纯函数无状态机） ｜ R7 N/A（无实例调用）
 * 修订历史 (Revision)   : 2026-11-20  v1.0.0  R50 首版（批次 1 · 序号 5）
 * 验收向量 (Acceptance) : ① 点 (0,0),(1,0),(0,1) → D=2.0，Ux=(0+1+0)/2=0.5，
 *                         Uy=(0+0+1)/2=0.5，R=SQRT(0.5)≈0.707106781186548，
 *                         返回 TRUE，eOk；② 点 (0,0),(1,1),(2,2) → D=2×
 *                         [0(1−2)+1(2−0)+2(0−1)]=0 → 共线拒绝，返回 FALSE，
 *                         eCollinear，三输出哨兵 0；③ x2=NaN → 返回 FALSE，
 *                         eNonFinite。
 *==============================================================================*)

(*-----------------------------------------------------------------------------
 * 枚举: E_DL_CircFitErr（错误码；故障级恒伴返回 FALSE）
 *----------------------------------------------------------------------------*)
TYPE E_DL_CircFitErr :
(
    eOk        := 0,   // 拟合成功 / Fit success
    eCollinear := 1,   // 故障级：三点共线（叉积绝对值低于容差） / Fault: three points collinear
    eNonFinite := 2    // 故障级：坐标非有限（NaN/Inf） / Fault: non-finite coordinate
);
END_TYPE

FUNCTION FC_DL_CircleFit3Pt : BOOL
VAR_INPUT
    fX1 : LREAL;                      // 点 1 横坐标 [mm] / Point 1 X coordinate [mm]
    fY1 : LREAL;                      // 点 1 纵坐标 [mm] / Point 1 Y coordinate [mm]
    fX2 : LREAL;                      // 点 2 横坐标 [mm] / Point 2 X coordinate [mm]
    fY2 : LREAL;                      // 点 2 纵坐标 [mm] / Point 2 Y coordinate [mm]
    fX3 : LREAL;                      // 点 3 横坐标 [mm] / Point 3 X coordinate [mm]
    fY3 : LREAL;                      // 点 3 纵坐标 [mm] / Point 3 Y coordinate [mm]
END_VAR
VAR_OUTPUT
    fCx      : LREAL;                 // 圆心横坐标（哨兵 0 于早退路径） [mm] / Centre X, sentinel zero on early exit [mm]
    fCy      : LREAL;                 // 圆心纵坐标 [mm] / Centre Y coordinate [mm]
    fR       : LREAL;                 // 外接圆半径 [mm] / Circumcircle radius [mm]
    eErrCode : E_DL_CircFitErr;       // 错误码出口 / Error code outlet
END_VAR
VAR
    _bNonFin : BOOL;                  // 六坐标非有限汇总 [-] / Non-finite aggregate flag
    _fD      : LREAL;                 // 行列式（2×叉积，除数） [mm²] / Determinant, 2 times cross product
    _fS1     : LREAL;                 // 点 1 平方和 x1²+y1² [mm²] / Point 1 squared norm
    _fS2     : LREAL;                 // 点 2 平方和 [mm²] / Point 2 squared norm
    _fS3     : LREAL;                 // 点 3 平方和 [mm²] / Point 3 squared norm
    _fUx     : LREAL;                 // 圆心横坐标中间量 [mm] / Centre X intermediate
    _fUy     : LREAL;                 // 圆心纵坐标中间量 [mm] / Centre Y intermediate
    _fDx     : LREAL;                 // 点 1 对圆心横差 [mm] / Point 1 to centre X difference
    _fDy     : LREAL;                 // 点 1 对圆心纵差 [mm] / Point 1 to centre Y difference
END_VAR
VAR CONSTANT
    DL_CFT_COLMIN : LREAL := 1.0E-9;  // 共线容差（|2×叉积| 低于此拒算，mm² 口径） [mm²] / Collinearity tolerance
    DL_CFT_ZERO   : LREAL := 0.0;     // 哨兵与非有限判零基准 [mm] / Sentinel and non-finite zero base
    DL_CFT_TWO    : LREAL := 2.0;     // 行列式系数 2 [-] / Determinant factor two
END_VAR

(* —— 段 0：出口预置安全值（四段式第一段：预置） —— *)
FC_DL_CircleFit3Pt := FALSE;          // 返回值预置无效 / Return preset invalid
fCx := DL_CFT_ZERO;                   // 圆心 X 哨兵 0 / Centre X sentinel
fCy := DL_CFT_ZERO;                   // 圆心 Y 哨兵 0 / Centre Y sentinel
fR := DL_CFT_ZERO;                    // 半径哨兵 0 / Radius sentinel
eErrCode := E_DL_CircFitErr.eNonFinite;   // 预置最严码 / Preset strictest code

(* —— 段 1：非有限域闸（R79 双判：NaN 自反 + Inf 差自减，六坐标逐一） —— *)
_bNonFin := (fX1 <> fX1) OR ((fX1 - fX1) <> DL_CFT_ZERO)
         OR (fY1 <> fY1) OR ((fY1 - fY1) <> DL_CFT_ZERO)
         OR (fX2 <> fX2) OR ((fX2 - fX2) <> DL_CFT_ZERO)
         OR (fY2 <> fY2) OR ((fY2 - fY2) <> DL_CFT_ZERO)
         OR (fX3 <> fX3) OR ((fX3 - fX3) <> DL_CFT_ZERO)
         OR (fY3 <> fY3) OR ((fY3 - fY3) <> DL_CFT_ZERO);   // 非有限汇总 / Non-finite aggregate
IF _bNonFin THEN
    RETURN;                           // 早退保持哨兵与最严码 / Early exit with sentinel
END_IF

(* —— 段 2：行列式与共线闸（D 作除数前置判，结构性无除零） —— *)
_fD := DL_CFT_TWO * (fX1 * (fY2 - fY3) + fX2 * (fY3 - fY1) + fX3 * (fY1 - fY2));   // D = 2×叉积 / Determinant
IF ABS(_fD) < DL_CFT_COLMIN THEN
    eErrCode := E_DL_CircFitErr.eCollinear;       // 共线拒绝（故障级，伴返回 FALSE） / Collinear reject
    RETURN;                                       // 早退保持哨兵 / Early exit with sentinel
END_IF

(* —— 段 3：代数内核（分母 D 已过闸） —— *)
_fS1 := fX1 * fX1 + fY1 * fY1;        // 点 1 平方和 / Point 1 squared norm
_fS2 := fX2 * fX2 + fY2 * fY2;        // 点 2 平方和 / Point 2 squared norm
_fS3 := fX3 * fX3 + fY3 * fY3;        // 点 3 平方和 / Point 3 squared norm
_fUx := (_fS1 * (fY2 - fY3) + _fS2 * (fY3 - fY1) + _fS3 * (fY1 - fY2)) / _fD;   // 圆心 X 解析解 / Centre X closed form
_fUy := (_fS1 * (fX3 - fX2) + _fS2 * (fX1 - fX3) + _fS3 * (fX2 - fX1)) / _fD;   // 圆心 Y 解析解 / Centre Y closed form
_fDx := fX1 - _fUx;                   // 点 1 对圆心横差 / X difference to centre
_fDy := fY1 - _fUy;                   // 点 1 对圆心纵差 / Y difference to centre

(* —— 段 4：半径合成与结果复检（平方和非负，无负开方；复检非有限兜底） —— *)
fR := SQRT(_fDx * _fDx + _fDy * _fDy);   // 半径 = 点 1 到圆心距离 / Radius via squared sum
IF (fR <> fR) OR ((fR - fR) <> DL_CFT_ZERO) THEN
    fCx := DL_CFT_ZERO;               // 复检异常回哨兵（四段式第四段） / Recheck failed: sentinel
    fCy := DL_CFT_ZERO;               // 回哨兵 / Sentinel
    fR := DL_CFT_ZERO;                // 回哨兵 / Sentinel
    RETURN;                           // 保持最严码早退 / Early exit strictest code
END_IF
fCx := _fUx;                          // 圆心 X 出口 / Centre X outlet
fCy := _fUy;                          // 圆心 Y 出口 / Centre Y outlet
eErrCode := E_DL_CircFitErr.eOk;      // 成功码 / Success code
FC_DL_CircleFit3Pt := TRUE;           // 拟合有效 / Fit valid

END_FUNCTION

(* ---- FC_DL_ConcentrationUnitConvert.st ---- *)
(*==============================================================================
 * 组件名称 (Component)  : FC_DL_ConcentrationUnitConvert
 * 所属子库 (Sublibrary) : DL_MathData
 * 当前版本 (Version)    : 1.0.0
 * 兼容性   (Platform)   : CODESYS 3.5+ / TwinCAT 3 / 汇川 InoProShop / 施耐德 Machine Expert
 *                         仅依赖 IEC 61131-3 算术运算符，零厂商私有库
 * 功能描述 (Function)   : 气体浓度单位换算：ppm（体积比）↔ %（体积比）↔ mg/m³（质量浓度）。
 *                         以 ppm 为中介单位：
 *                           %      → ppm   : × 10000
 *                           mg/m3  → ppm   : × Vm / M           （Vm = 22.414 L/mol）
 *                           ppm    → mg/m3 : × M / Vm
 *                         **标况假设（显式声明）**：Vm = 22.414 L/mol 为 0 ℃、101.325 kPa
 *                         干气理想气体摩尔体积；本件不做温压修正，非标况数据必须先由调用方
 *                         折算至标况再调用本件。摩尔质量 M 由引脚传入（g/mol），
 *                         不同气体（CO / CH4 / VOC 等）必须分别给值。
 * 接口     (Interface)  : 输入 fValue 被换算浓度 [源单位]、eSrc 源单位、eDst 目标单位、
 *                         fMolarMass 摩尔质量 [g/mol]（**换算必需，必须 > 0**）；
 *                         输出 fConverted 换算结果 [目标单位]、eErrCode（E_DL_ConcConvErr）；
 *                         返回值 = bValid 数值可信标志（TRUE = fConverted 可信）。
 * 边界     (Boundary)   : ① 属主边界：只做单位换算，不做温压折算、不做多组分加权、不做报警阈值比较。
 *                         ② **除零防护（R4 硬要求）**：mg/m³ ↔ ppm 两个方向都含除以 M 或除以 Vm 的
 *                         路径，进入分支前先判 fMolarMass > 0，否则故障级 eInvalidMolarMass 早退。
 *                         ③ 全部浮点入参非有限双判（fValue 与 fMolarMass 逐一枚举）。
 *                         ④ 浓度非负：负值 → 故障级 eNegativeValue（浓度无负值语义）。
 *                         ⑤ 单位枚举越域 → 故障级 eInvalidUnit，结果哨兵 0。
 *                         ⑥ ppm 与 % 为体积比，其换算不依赖 M；mg/m³ 参与的两向换算才依赖 M。
 *                         ⑦ 零全局耦合（无 GVL / VAR_EXTERNAL / 物理地址）。
 * 分工声明 (Scope)      : 与 `FC_DL_HumidityUnitConvert` 分工：湿度归那件；
 *                         与气体检测 FB（未入库）分工：报警分级与延时归那件，本件只换算数值。
 * 来源标签 (Source Tag) : 开源溯源：lgf-math 换算系数（公开物理常数，clean-room 重写）；许可证 MIT（仅参考语义，代码原创）
 * 码表     (Codes)      : 本件不占用全局数字码位；出口为 BOOL + LREAL +
 *                         本文件内定义 enum E_DL_ConcConvErr（全库唯一）。
 * 红线自检 (Redline)    : R1 ✓ 零 GVL/VAR_EXTERNAL ｜ R2 ✓ 零 %I/%Q/%M ｜ R3 ✓ 纯 IEC 61131-3
 *                         R4 ✓ 摩尔质量前置判零 + 全浮点非有限双判 + 负值拒绝 ｜ R5 ✓ 声明逐行同行双语注释
 *                         R6 N/A（纯函数无状态机） ｜ R7 N/A（无实例调用）
 * 修订历史 (Revision)   : 2026-11-23  v1.0.0  R77 首版（批次 B2 · 序号 20）
 * 验收向量 (Acceptance) : ① fValue=1.0(%) , eSrc=ePercent, eDst=ePpm → 1×10000 = 10000.0 ppm, eOk, TRUE；
 *                         ② fValue=10000.0, eSrc=ePpm, eDst=ePercent → 1.0 %, eOk；
 *                         ③ fValue=100.0(mg/m3), eSrc=eMgM3, eDst=ePpm, fMolarMass=28.01(CO) →
 *                         100×22.414/28.01 ≈ 80.0214 ppm（容差 1E-3）；
 *                         ④ fValue=80.0214, eSrc=ePpm, eDst=eMgM3, fMolarMass=28.01 →
 *                         80.0214×28.01/22.414 ≈ 100.0 mg/m3（容差 1E-2，与 ③ 互逆）；
 *                         ⑤ fMolarMass=0.0 → 返回 FALSE, 0, eInvalidMolarMass（除零防护分支）；
 *                         ⑥ fValue=-1.0, eSrc=ePpm, eDst=ePercent → 返回 FALSE, 0, eNegativeValue。
 *==============================================================================*)

(*-----------------------------------------------------------------------------
 * 枚举: E_DL_ConcUnit（气体浓度单位表，归属 DL_MathData，与本件同文件，全库唯一属主）
 *----------------------------------------------------------------------------*)
TYPE E_DL_ConcUnit :
(
    ePpm     := 0,   // 百万分之一（体积比，中介单位） / Parts per million by volume, hub unit
    ePercent := 1,   // 体积百分数（= 10000 ppm） / Volume percent
    eMgM3    := 2    // 毫克每立方米（质量浓度，需摩尔质量换算） / Milligrams per cubic metre, needs molar mass
);
END_TYPE

(*-----------------------------------------------------------------------------
 * 枚举: E_DL_ConcConvErr（浓度换算错误码）
 *----------------------------------------------------------------------------*)
TYPE E_DL_ConcConvErr :
(
    eOk               := 0,   // 信息级：换算完成 / Info: conversion completed
    eZeroValue        := 1,   // 信息级：输入为零（合法） / Info: zero input, legal
    eInvalidUnit      := 2,   // 故障级：单位枚举越域 / Fault: unit enum out of domain
    eNonFinite        := 3,   // 故障级：入参非有限 / Fault: non-finite input
    eNegativeValue    := 4,   // 故障级：负浓度 / Fault: negative concentration
    eInvalidMolarMass := 5    // 故障级：摩尔质量非正，除零风险 / Fault: molar mass not positive, division-by-zero risk
);
END_TYPE

FUNCTION FC_DL_ConcentrationUnitConvert : BOOL
VAR_INPUT
    fValue     : LREAL;         // 被换算浓度值 [源单位] / Concentration value in source unit
    eSrc       : E_DL_ConcUnit; // 源单位枚举 [-] / Source unit enum
    eDst       : E_DL_ConcUnit; // 目标单位枚举 [-] / Destination unit enum
    fMolarMass : LREAL;         // 摩尔质量（换算必需，必须 > 0） [g/mol] / Molar mass, mandatory and positive [g/mol]
END_VAR
VAR_OUTPUT
    fConverted : LREAL;             // 换算结果 [目标单位] / Converted result
    eErrCode   : E_DL_ConcConvErr;  // 错误码出口 [-] / Error code outlet
END_VAR
VAR
    _bNonFin : BOOL;   // 入参非有限当拍标志 [-] / Non-finite input flag
    _bNeedMol: BOOL;   // 本次换算是否需要摩尔质量 [-] / Whether molar mass is used in this conversion
    _fHub    : LREAL;  // 中介浓度值 [ppm] / Hub concentration value in ppm
END_VAR
VAR CONSTANT
    DL_CUC_PCT   : LREAL := 10000.0;   // % → ppm 换算系数（1% = 10000 ppm） [-] / Percent to ppm factor
    DL_CUC_VM    : LREAL := 22.414;    // 标况摩尔体积（0 ℃, 101.325 kPa） [L/mol] / Molar volume at standard conditions
    DL_CUC_ONE   : LREAL := 1.0;       // ppm 恒等系数 [-] / ppm identity factor
    DL_CUC_ZERO  : LREAL := 0.0;       // 零基准与非有限判零基准 [-] / Zero and non-finite base
    DL_CUC_TINY  : LREAL := 1.0E-9;    // 参数近似零阈值 [g/mol] / Near-zero parameter threshold
END_VAR

(* —— 段 0：出口预置安全值 —— *)
FC_DL_ConcentrationUnitConvert := FALSE;           // 返回值预置无效 / Return preset invalid
fConverted := DL_CUC_ZERO;                         // 结果哨兵 0 / Result sentinel
eErrCode   := E_DL_ConcConvErr.eInvalidUnit;       // 预置最严码 / Preset strictest code

(* —— 段 1：非有限域闸（fValue 与 fMolarMass 逐一枚举，禁止漏闸） —— *)
_bNonFin := (fValue <> fValue) OR ((fValue - fValue) <> DL_CUC_ZERO);            // 浓度值非有限 / Concentration non-finite
_bNonFin := _bNonFin OR (fMolarMass <> fMolarMass) OR ((fMolarMass - fMolarMass) <> DL_CUC_ZERO);  // 摩尔质量非有限 / Molar mass non-finite
IF _bNonFin THEN
    eErrCode := E_DL_ConcConvErr.eNonFinite;       // 故障级码 / Fault-level code
    RETURN;
END_IF

(* —— 段 2：单位枚举域闸 —— *)
IF (eSrc <> E_DL_ConcUnit.ePpm) AND (eSrc <> E_DL_ConcUnit.ePercent) AND (eSrc <> E_DL_ConcUnit.eMgM3) THEN
    RETURN;                                        // 源单位越域 / Source unit out of domain
END_IF
IF (eDst <> E_DL_ConcUnit.ePpm) AND (eDst <> E_DL_ConcUnit.ePercent) AND (eDst <> E_DL_ConcUnit.eMgM3) THEN
    RETURN;                                        // 目标单位越域 / Destination unit out of domain
END_IF

(* —— 段 3：负浓度域闸 —— *)
IF fValue < DL_CUC_ZERO THEN
    eErrCode := E_DL_ConcConvErr.eNegativeValue;   // 故障级码 / Fault-level code
    RETURN;
END_IF

(* —— 段 4：摩尔质量前置判零（凡涉及 mg/m3 的换算方向都必须先过此闸） —— *)
_bNeedMol := (eSrc = E_DL_ConcUnit.eMgM3) OR (eDst = E_DL_ConcUnit.eMgM3);   // 是否需要摩尔质量 / Molar mass needed flag
IF _bNeedMol THEN
    IF fMolarMass < DL_CUC_TINY THEN
        eErrCode := E_DL_ConcConvErr.eInvalidMolarMass;   // 故障级：摩尔质量非正 / Fault: non-positive molar mass
        RETURN;                                            // 早退，杜绝除以非正量 / Early exit, avoids division by non-positive value
    END_IF
END_IF

(* —— 段 5：源单位 → 中介 ppm —— *)
IF eSrc = E_DL_ConcUnit.ePpm THEN
    _fHub := fValue * DL_CUC_ONE;                  // ppm 直通 / ppm pass-through
ELSIF eSrc = E_DL_ConcUnit.ePercent THEN
    _fHub := fValue * DL_CUC_PCT;                  // % × 10000 / Percent scaled
ELSE
    _fHub := fValue * DL_CUC_VM / fMolarMass;      // mg/m3 × Vm / M（M 已在段 4 判正） / Mass to volume ppm
END_IF

(* —— 段 6：中介 ppm → 目标单位 —— *)
IF eDst = E_DL_ConcUnit.ePpm THEN
    fConverted := _fHub / DL_CUC_ONE;              // ÷1 直通 / Divide by identity
ELSIF eDst = E_DL_ConcUnit.ePercent THEN
    fConverted := _fHub / DL_CUC_PCT;              // ÷10000 / Divide by percent factor
ELSE
    fConverted := _fHub * fMolarMass / DL_CUC_VM;  // ppm × M / Vm（Vm 为常量 22.414，M 已判正） / Volume to mass
END_IF

(* —— 段 7：结果非有限复检兜底 —— *)
IF (fConverted <> fConverted) OR ((fConverted - fConverted) <> DL_CUC_ZERO) THEN
    fConverted := DL_CUC_ZERO;                     // 复检异常回哨兵 / Recheck failed: sentinel
    eErrCode   := E_DL_ConcConvErr.eNonFinite;     // 故障级码 / Fault-level code
    RETURN;
END_IF

(* —— 段 8：成功出口 —— *)
IF fValue = DL_CUC_ZERO THEN
    eErrCode := E_DL_ConcConvErr.eZeroValue;       // 信息级：零值 / Info: zero value
ELSE
    eErrCode := E_DL_ConcConvErr.eOk;              // 信息级成功 / Info success
END_IF
FC_DL_ConcentrationUnitConvert := TRUE;            // 换算有效 / Conversion valid

END_FUNCTION

(* ---- FC_DL_CovarOnline.st ---- *)
(*==============================================================================
 * 组件名称 (Component)  : FC_DL_CovarOnline
 * 所属子库 (Sublibrary) : DL_MathData
 * 当前版本 (Version)    : 1.0.0
 * 兼容性   (Platform)   : CODESYS 3.5+ / TwinCAT 3 / 汇川 InoProShop / 施耐德 Machine Expert
 *                         仅依赖 IEC 61131-3 基本算术，零厂商私有库
 * 功能描述 (Function)   : 双信号在线协方差（Welford 增量式），单遍流式更新、免二次遍历。
 *                         每拍只吃一对样本 (fX, fY)，把状态推进到调用者持有的累加结构 ST_DL_CovarAcc 中，
 *                         因此"在线"语义靠 IN_OUT 携带状态实现，函数本体无隐式记忆量。
 *                         Welford 协方差增量式（与均值更新交替，数值稳定）：
 *                           n ← n + 1                       （先计数，n 恒 ≥ 1）
 *                           dx ← x − meanX                  （用旧均值）
 *                           meanX ← meanX + dx / n
 *                           dy ← y − meanY
 *                           meanY ← meanY + dy / n
 *                           C ← C + dx · (y − meanY)        （用**新**均值，cosvar 更新式）
 *                           协方差 = C / (n − 1)            （样本协方差，n ≥ 2 才有定义）
 *                         验收向量（退化为可解析预测，R105 退化自检）：
 *                           ① 三点共线 y = 2x（x=1,2,3）→ 协方差 = 4.0，方差域比 = 1
 *                           ② 常量序列 x≡y≡5（n≥2）      → 协方差 = 0.0（差值容差内）
 *                           ③ 单样本 n=1                  → bValid=FALSE，不宣称
 * 接口     (Interface)  : IN_OUT stAcc 累加体（n/meanX/meanY/C 四量，调用者持有并负责复位）；
 *                         入 fX 样本 X、fY 样本 Y；出 返回值 = 样本协方差、bValid 宣称位（n≥2）、
 *                         bSampleRejected 当拍样本被剔标志、bResetDone 首样本生效标志。
 * 边界     (Boundary)   : ① **非有限样本前置剔除**：任一路为 NaN（自反判定 x<>x）或 Inf
 *                         （差值自反 (x−x)<>(x−x)）→ 当拍不累加、返回上一次已算协方差、置
 *                         bSampleRejected；② **分母闸**：n<2 时不做除法，返回 0 + bValid=FALSE
 *                         （单样本协方差无定义，绝不能拿 0/0 出来）；③ **输出钳位**：
 *                         协方差绝对值超 fCovarMax 时钳到 ±fCovarMax（防上游 IEEE 单位换算爆表）；
 *                         ④ 浮点比较一律差值容差，禁 = / <>（本件仅在 ABS 差 < 1E-12 处判等）；
 *                         ⑤ 累加体越界（n 达 UDINT 上限）时整体冻结不再累加并置 bSampleRejected；
 *                         ⑥ 零全局耦合、零物理地址。
 * 分工声明 (Scope)      : 本件只做"双流协方差原子件"。不接管：单信号多统计量聚合
 *                         （属 FB_DL_SignalStatistics）、相关系数归一（由调用者自行除以 σx·σy）、
 *                         样本窗口滑窗淘汰（本件是全历史累加，滑窗属上层窗口件）。
 * 来源标签 (Source Tag) : T2-1 LGF · Measurement ◐（流式协方差，自研 clean-room）
 * 码表     (Codes)      : 本件不占用任何全局数字码位（零码位范式 R297）；诊断由 BOOL 出口承担。
 * 红线自检 (Redline)    : R1 ✓ 零 GVL/VAR_EXTERNAL ｜ R2 ✓ 零 %I/%Q/%M ｜ R3 ✓ 纯 IEC 61131-3
 *                         R4 ✓ 非有限剔除 + 分母闸 + 输出钳位 + 差值容差 ｜ R5 ✓ 声明逐行同行双语注释
 *                         R6 ✓ 无状态机（纯组合函数，判别 IF 链带兜底分支） ｜ R7 ✓ 无定时器/沿实例
 * 修订历史 (Revision)   : 2026-11-19  v1.0.0  R47 首版（批次 1 · 序号 3）
 *==============================================================================*)

TYPE ST_DL_CovarAcc :
STRUCT
    nCnt  : UDINT := 0;     // 已收样本数（含当拍） [个] / Accepted sample count including this scan
    fMeanX: LREAL := 0.0;   // X 流运行均值 [工程单位] / Running mean of the X stream
    fMeanY: LREAL := 0.0;   // Y 流运行均值 [工程单位] / Running mean of the Y stream
    fC    : LREAL := 0.0;   // 协方差分子累加量 C = Σ(x−mx)(y−my) [单位²] / Covariance co-moment accumulator
    fLast : LREAL := 0.0;   // 上次有效协方差（被剔样本当拍回放） [单位²] / Last valid covariance, replayed on reject
END_STRUCT
END_TYPE

FUNCTION FC_DL_CovarOnline : LREAL
VAR_IN_OUT
    stAcc : ST_DL_CovarAcc;                 // 累加体（调用者持有；复位时四量清 0） [-] / Accumulator owned by the caller
END_VAR
VAR_INPUT
    fX        : LREAL := 0.0;               // X 流当拍样本 [工程单位] / X sample of this scan
    fY        : LREAL := 0.0;               // Y 流当拍样本 [工程单位] / Y sample of this scan
    fCovarMax : LREAL := 1.0E12;            // 协方差输出绝对上限，域 > 0 [单位²] / Absolute covariance clamp, > 0
END_VAR
VAR_OUTPUT
    bValid          : BOOL := FALSE;        // 宣称位（n≥2 且本次除法合法） [-] / Validity flag, n >= 2
    bSampleRejected : BOOL := FALSE;        // 当拍样本被剔（非有限或计数饱和） [-] / Sample rejected this scan
END_VAR
VAR
    bXFin : BOOL := FALSE;                  // X 样本有限性判定中间量 [-] / X finiteness working flag
    bYFin : BOOL := FALSE;                  // Y 样本有限性判定中间量 [-] / Y finiteness working flag
    fDx   : LREAL := 0.0;                   // X 相对旧均值偏差 [工程单位] / X deviation from the old mean
    fDy   : LREAL := 0.0;                   // Y 相对旧均值偏差 [工程单位] / Y deviation from the old mean
    fN    : LREAL := 0.0;                   // 样本数的实数副本（作除数，已证 ≥ 1） [-] / Real copy of the count
    fLim  : LREAL := 0.0;                   // 生效钳位限（脚非法时回退常量，R127 解耦） [单位²] / Effective clamp limit
    fOut  : LREAL := 0.0;                   // 结果工作值 [单位²] / Result working value
END_VAR
VAR CONSTANT
    DL_COV_LIM_DEF : LREAL := 1.0E12;       // 钳位限回退默认值（与脚默认同源） [单位²] / Default clamp limit
    DL_COV_CNT_MAX : UDINT := 16#FFFF_FFFE; // 样本计数饱和闸（留 1 个余量防 +1 回绕） [个] / Count saturation gate
    DL_COV_EPS     : LREAL := 1.0E-12;      // 浮点判等容差（仅用于"差≈0"判定） [-] / Equality tolerance
END_VAR

(* —— 段 1：返回值与标志预置（R45 四段式第①段） —— *)
FC_DL_CovarOnline := 0.0;                   // 返回值预置 / Return value preset
bValid := FALSE;                            // 宣称位预置 / Validity preset
bSampleRejected := FALSE;                   // 剔除标志预置 / Reject flag preset
fOut := 0.0;                                 // 结果工作值预置 / Result working preset

(* —— 段 2：钳位限域闸（脚值非法回退常量，二级钳定 R117；R127 兜底值与被判量解耦） —— *)
fLim := fCovarMax;                           // 先直取脚值 / Take the pin value first
IF (fLim <> fLim) OR ((fLim - fLim) <> (fLim - fLim)) OR (fLim <= 0.0) THEN
    fLim := DL_COV_LIM_DEF;                  // 非有限或非正：回退默认常量 / Non-finite or non-positive: fall back
END_IF

(* —— 段 3：样本有限性闸（NaN 自反 + Inf 差值自反，LREAL 域无幅值常量可用，R40） —— *)
bXFin := NOT ((fX <> fX) OR ((fX - fX) <> (fX - fX)));      // X 有限 ⇔ 非 NaN 且非 Inf / X finite
bYFin := NOT ((fY <> fY) OR ((fY - fY) <> (fY - fY)));      // Y 有限 ⇔ 非 NaN 且非 Inf / Y finite

(* —— 段 4：剔除分支（非有限或计数饱和：不累加，回放上次有效值） —— *)
IF (NOT bXFin) OR (NOT bYFin) OR (stAcc.nCnt >= DL_COV_CNT_MAX) THEN
    bSampleRejected := TRUE;                 // 当拍样本拒收 / Reject this scan's sample
    fOut := stAcc.fLast;                     // 回放上次有效协方差（保持槽非有限闸已在写入侧保证） / Replay last valid value
ELSE
    (* —— 段 5：Welford 增量更新（先计数，再双均值，最后共矩） —— *)
    stAcc.nCnt := stAcc.nCnt + 1;            // 计数先推进（n ≥ 1，除零结构性不可能） / Count first, n >= 1 guaranteed
    fN := UDINT_TO_LREAL(stAcc.nCnt);        // 实数副本作除数 / Real copy as divisor

    fDx := fX - stAcc.fMeanX;                // X 偏差（旧均值） / X deviation from old mean
    stAcc.fMeanX := stAcc.fMeanX + (fDx / fN);   // X 均值更新 / Update X mean
    fDy := fY - stAcc.fMeanY;                // Y 偏差（旧均值） / Y deviation from old mean
    stAcc.fMeanY := stAcc.fMeanY + (fDy / fN);   // Y 均值更新 / Update Y mean

    stAcc.fC := stAcc.fC + (fDx * (fY - stAcc.fMeanY));  // 共矩增量（用新均值） / Co-moment increment with the new mean

    IF stAcc.nCnt >= 2 THEN
        fOut := stAcc.fC / (fN - 1.0);       // 样本协方差（分母 n−1 ≥ 1） / Sample covariance
        bValid := TRUE;                       // 样本数够：允许宣称 / Enough samples: may claim validity
    ELSE
        fOut := 0.0;                          // 单样本：协方差无定义，输出 0 / Single sample: undefined, output 0
        bValid := FALSE;                      // 不宣称 / Do not claim
    END_IF
END_IF

(* —— 段 6：结果非有限复检 + 钳位（R45 四段式第④段） —— *)
IF (fOut <> fOut) OR ((fOut - fOut) <> (fOut - fOut)) THEN
    fOut := 0.0;                             // 结果非有限：归 0 / Non-finite result: zeroed
    bValid := FALSE;                          // 同步撤宣称 / Withdraw validity in the same scan
END_IF
IF fOut > fLim THEN
    fOut := fLim;                             // 上钳 / Clamp high
ELSIF fOut < (0.0 - fLim) THEN
    fOut := 0.0 - fLim;                       // 下钳（写作 0.0−lim，避免负号字面量歧义） / Clamp low
END_IF

(* —— 段 7：保持槽写入（仅有限值可写入信任根，R133） —— *)
IF (NOT bSampleRejected) AND bValid THEN
    stAcc.fLast := fOut;                      // 记录最近有效值 / Remember the latest valid value
END_IF

(* —— 段 8：统一出口 —— *)
FC_DL_CovarOnline := fOut;                    // 输出样本协方差 / Output the sample covariance

END_FUNCTION

(* ---- FC_DL_Crc16Ccitt.st ---- *)
(*
    FC_DL_Crc16Ccitt —— CRC-16 三变体位算法（多项式 0x1021 族）
    ------------------------------------------------------------------
    分类      : DL_MathData / Checksum
    前缀      : FC_DL_
    版本      : 1.0.1
    溯源      : T2-1 LGF · Data Handling（源矩阵明列「校验族尚余 CRC-16 反射待挖」）；
                T1-3 OSCAT Network 校验族分类为次源，不复制实现；
                参数集与校验值经一次公开资料核对（三家在线 CRC 计算器一致）；
                clean-room 重写，未复制任何闭源厂商源码，参考实现仅限 MIT/Apache 许可
    平台      : 纯 IEC 61131-3，CODESYS V3.5+ / TwinCAT 3 / InoProShop 通用
    作者      : 道莅代码库 · PLC编程专家（R18）
    ------------------------------------------------------------------
    功能说明  : 一个函数覆盖 CRC-16 三个最常用参数集（同一多项式 0x1021 的三种参数化），
                解决现场「设备手册只写 CRC-16 CCITT，不说 init / 反射」导致的对接失败；
                库内 FC_DL_Crc16Modbus 已占 0x8005 反射族，本件补 0x1021 族；
                反射变体不使用任何位反指令（跨平台可用性风险），改用「右移 + 判最低位」
                循环实现，三个变体共用同一份位循环骨架；
                位循环定长 8 次，无 WHILE，循环次数可静态界定。
    验收向量  : 对 "123456789"（9 字节）逐字节调用后应得
                eCrc16CcittFalse = 16#29B1 ｜ eCrc16Xmodem = 16#31C3 ｜ eCrc16Kermit = 16#2189
    错误码    : 16#0001_023D uLen 超 256 已截断，仅校验前 256 字节——信息级，正常防御
                16#0001_023E 预留禁用（信息级，不得挪用）
                16#0001_0312 预留禁用（故障级，不得挪用；空帧非法方言的预留归属，实现体内零赋值）
                16#0001_0313 变体枚举值非法（CASE 落 ELSE）——故障级，返回 0
                16#0001_0314 预留禁用（故障级，不得挪用）
    码位总账  : 16#0001_023D 用 / 16#0001_023E 预留 ｜ 16#0001_0312 预留 / 16#0001_0313 用 / 16#0001_0314 预留
    状态机    : N/A —— 纯函数无顺序状态机，无 CASE 可写（变体枚举选择用 CASE 且含 ELSE 兜底）
    采样约定  : 纯组合函数，无定时器、无内部驻留状态；uLen = 0 为空帧，返回 init 值且 bValid 为 TRUE，
                空帧是协议合法输入，不按故障处理。
    修订记录  : 2026-11-16 v1.0.0 首次入库（R18）
                2026-11-16 v1.0.1 R18 终审修复：uLen = 0 时 FOR 终止表达式 uLenEff - 1 在 UINT 下回绕成
                65535，越界读 auData[256..65535] 触发运行时数组越界；改为空帧短路提前返回 init 值，
                循环段保证 uLenEff >= 1。对外引脚与校验值零变更。
*)

(*-----------------------------------------------------------------------------
 * 枚举: E_DL_Crc16Vari（归属本函数，与其同文件发布）
 * 含义: CRC-16 参数集选择，成员值写死便于工程持久化
 *----------------------------------------------------------------------------*)
TYPE E_DL_Crc16Vari :
(
    eCrc16CcittFalse := 0,   // CCITT-FALSE：poly 0x1021 / init 0xFFFF / 不反射 / 无终值异或 / CCITT-FALSE, init 0xFFFF, no reflection, no final xor
    eCrc16Xmodem     := 1,   // XMODEM：poly 0x1021 / init 0x0000 / 不反射 / 无终值异或 / XMODEM, init 0x0000, no reflection, no final xor
    eCrc16Kermit     := 2    // KERMIT：poly 0x8408（位反形式）/ init 0x0000 / 入出均反射 / KERMIT, reflected poly 0x8408, init 0x0000, reflected in and out
) UINT;
END_TYPE

FUNCTION FC_DL_Crc16Ccitt : WORD
VAR_INPUT
    auData : ARRAY[0..255] OF BYTE;                          // 待校验字节数组，定长 256，超长由 uLen 截断 [字节] / data bytes, fixed length 256, truncated by uLen [byte]
    uLen   : UINT := 0;                                      // 有效长度 [字节]，范围 0~256，0 = 空帧 / valid length [byte], range 0~256, 0 = empty frame
    eVari  : E_DL_Crc16Vari := E_DL_Crc16Vari.eCrc16CcittFalse; // 参数集选择 / parameter set selection
END_VAR
VAR_OUTPUT
    eErr   : UDINT;                                          // 错误码，0=正常 / error id, 0=ok
    bError : BOOL;                                           // 故障标志，eErr 为故障级时 TRUE / error flag, TRUE on fault-level eErr
    bValid : BOOL;                                           // 结果是否可用，故障态 FALSE / result usable flag, FALSE in fault state
END_VAR
VAR
    uCrc     : WORD;                                         // CRC 寄存器 [无量纲] / CRC register [dimensionless]
    uPoly    : WORD;                                         // 生效多项式，由变体决定 [无量纲] / active polynomial selected by the variant [dimensionless]
    uIdx     : UINT;                                         // 字节游标 [字节] / byte cursor [byte]
    nBit     : INT;                                          // 位游标 0~7 [位] / bit cursor 0~7 [bit]
    uByte    : BYTE;                                         // 当前处理字节 [字节] / byte under processing [byte]
    bReflect : BOOL;                                         // 反射变体标志，TRUE 走右移分支 / reflected variant flag, TRUE takes the right-shift branch
    uLenEff  : UINT;                                         // 生效长度，截断后使用 [字节] / effective length after truncation [byte]
END_VAR
VAR CONSTANT
    DL_CRC16_LEN_MAX     : UINT := 256;                      // 长度上限 [字节] / length upper bound [byte]
    DL_CRC16_POLY_MSB    : WORD := 16#1021;                  // 高位先行多项式 [无量纲] / most significant bit first polynomial [dimensionless]
    DL_CRC16_POLY_LSB    : WORD := 16#8408;                  // 低位先行（位反）多项式 [无量纲] / least significant bit first (reflected) polynomial [dimensionless]
    DL_CRC16_INIT_FFFF   : WORD := 16#FFFF;                  // 全一初值 [无量纲] / all ones initial value [dimensionless]
    DL_CRC16_INIT_ZERO   : WORD := 16#0000;                  // 全零初值 [无量纲] / all zeros initial value [dimensionless]
    DL_CRC16_BIT_MSB     : WORD := 16#8000;                  // 最高位掩码 [位图] / most significant bit mask [bitmap]
    DL_CRC16_BIT_LSB     : WORD := 16#0001;                  // 最低位掩码 [位图] / least significant bit mask [bitmap]
    DL_CRC16_SHIFT_BYTE  : INT := 8;                         // 字节位宽，左移量恒为 8 [位] / byte width, the left shift is always 8 [bit]
    DL_CRC16_BIT_LAST    : INT := 7;                         // 位循环末值 [位] / last index of the bit loop [bit]
    DL_CRC16_LEN_NONE    : UINT := 0;                        // 空帧长度哨兵，用于 UINT 减法前判零 [字节] / empty frame length sentinel, guards the UINT subtraction [byte]
    DL_CRC16_CHECK_CCITT : WORD := 16#29B1;                  // "123456789" 的 CCITT-FALSE 校验值（验收向量）[无量纲] / check value for "123456789", CCITT-FALSE [dimensionless]
    DL_CRC16_CHECK_XMODEM: WORD := 16#31C3;                  // "123456789" 的 XMODEM 校验值（验收向量）[无量纲] / check value for "123456789", XMODEM [dimensionless]
    DL_CRC16_CHECK_KERMIT: WORD := 16#2189;                  // "123456789" 的 KERMIT 校验值（验收向量）[无量纲] / check value for "123456789", KERMIT [dimensionless]
END_VAR

// 段 1｜返回值与错误状态预置 / segment 1, preset return value and error status
FC_DL_Crc16Ccitt := DL_CRC16_INIT_ZERO;        // 故障缺省返回 0 / fault default returns zero
eErr := 0;                                     // 预置无错误 / preset no error
bError := FALSE;                               // 预置无故障 / preset no fault
bValid := FALSE;                               // 预置结果不可用，通过闸门后置位 / preset unusable, set TRUE after the gates
uLenEff := uLen;                               // 默认沿用输入长度 / default to the input length

// 段 2｜长度闸：超上限先截断再校验，绝不越界读 / segment 2, length gate truncates before any read
IF uLen > DL_CRC16_LEN_MAX THEN
    uLenEff := DL_CRC16_LEN_MAX;               // 截断到 256 字节 / truncate to 256 bytes
    eErr := 16#0001_023D;                      // 截断提示（信息级不置故障）/ truncation hint, info level never raises a fault
END_IF

// 段 3｜变体参数装载（CASE 必须含 ELSE 兜底，红线）/ segment 3, load the variant parameters
CASE eVari OF
    E_DL_Crc16Vari.eCrc16CcittFalse :
        uCrc := DL_CRC16_INIT_FFFF;            // 全一初值 / all ones initial value
        uPoly := DL_CRC16_POLY_MSB;            // 高位先行多项式 / most significant bit first polynomial
        bReflect := FALSE;                     // 不反射 / no reflection
    E_DL_Crc16Vari.eCrc16Xmodem :
        uCrc := DL_CRC16_INIT_ZERO;            // 全零初值 / all zeros initial value
        uPoly := DL_CRC16_POLY_MSB;            // 高位先行多项式 / most significant bit first polynomial
        bReflect := FALSE;                     // 不反射 / no reflection
    E_DL_Crc16Vari.eCrc16Kermit :
        uCrc := DL_CRC16_INIT_ZERO;            // 全零初值 / all zeros initial value
        uPoly := DL_CRC16_POLY_LSB;            // 位反多项式 / reflected polynomial
        bReflect := TRUE;                      // 入出均反射 / reflected in and out
ELSE
    eErr := 16#0001_0313;                      // 变体枚举非法故障码 / illegal variant enum fault id
    bError := TRUE;                            // 置故障标志 / raise the error flag
    bValid := FALSE;                           // 结果不可用 / result unusable
    FC_DL_Crc16Ccitt := DL_CRC16_INIT_ZERO;    // 返回 0 / return zero
    RETURN;                                    // 故障级提前返回 / early return on fault
END_CASE

// 段 4｜空帧短路：UINT 下 uLenEff - 1 在 uLenEff = 0 时回绕成 65535，直接进循环会越界读 / segment 4, empty frame short circuit
// 说明：IEC 61131-3 的 FOR 终止表达式在进入循环时求值一次，故 0 - 1 必然回绕，必须先判零再做减法
IF uLenEff = DL_CRC16_LEN_NONE THEN
    FC_DL_Crc16Ccitt := uCrc;                  // 空帧返回 init 值 / an empty frame returns the initial value
    bValid := TRUE;                            // 空帧是协议合法输入 / an empty frame is a legal protocol input
    RETURN;                                    // 提前出口，绝不进循环 / early exit, never enter the loop
END_IF

// 段 4b｜逐字节位算法：uLenEff 已保证 >= 1，减法安全 / segment 4b, byte by byte bit algorithm with a safe subtraction
FOR uIdx := 0 TO uLenEff - 1 DO
    uByte := auData[uIdx];                     // 取当前字节，索引上界已由长度闸保证 / fetch the byte, the upper bound is guaranteed by the length gate
    IF bReflect THEN
        uCrc := uCrc XOR BYTE_TO_WORD(uByte);  // 反射变体：低字节对齐异或 / reflected variant, low byte aligned xor
        FOR nBit := 0 TO DL_CRC16_BIT_LAST DO
            IF (uCrc AND DL_CRC16_BIT_LSB) <> 0 THEN
                uCrc := SHR(uCrc, 1) XOR uPoly; // 最低位为 1 则右移后异或多项式 / shift right and xor the polynomial when the lowest bit is set
            ELSE
                uCrc := SHR(uCrc, 1);          // 最低位为 0 只右移 / shift right only when the lowest bit is clear
            END_IF
        END_FOR
    ELSE
        uCrc := uCrc XOR SHL(BYTE_TO_WORD(uByte), DL_CRC16_SHIFT_BYTE); // 高位先行：字节左移 8 位异或 / msb first, xor the byte shifted left by eight
        FOR nBit := 0 TO DL_CRC16_BIT_LAST DO
            IF (uCrc AND DL_CRC16_BIT_MSB) <> 0 THEN
                uCrc := SHL(uCrc, 1) XOR uPoly; // 最高位为 1 则左移后异或多项式 / shift left and xor the polynomial when the highest bit is set
            ELSE
                uCrc := SHL(uCrc, 1);          // 最高位为 0 只左移 / shift left only when the highest bit is clear
            END_IF
        END_FOR
    END_IF
END_FOR

// 段 5｜出口：空帧是协议合法输入，bValid 仍为 TRUE / segment 5, exit, an empty frame is a legal protocol input
FC_DL_Crc16Ccitt := uCrc;                      // 输出寄存器值 / publish the register value
bValid := TRUE;                                // 结果可用 / the result is usable
END_FUNCTION

(* ---- FC_DL_DeltaClampReal.st ---- *)
(*==============================================================================
 * 组件名称 (Component)  : FC_DL_DeltaClampReal
 * 所属子库 (Sublibrary) : DL_MathData ｜ 版本 (Version) : 1.0.0 ｜ 2026-11-23
 * 兼容性   (Platform)   : CODESYS 3.5+ / TwinCAT 3 / 汇川 InoProShop / 施耐德 Machine Expert
 *                         仅依赖 IEC 61131-3 算术运算符与 ABS，零厂商私有库
 * 功能描述 (Function)   : 相邻两拍增量钳位（FC 形态）：|fX − fXPrev| 超过 fMaxDelta 时，
 *                         输出改为 fXPrev 沿增量方向叠加 fMaxDelta（钳位后叠加，非就地截断），
 *                         未超限则直通 fX。用于抑制单拍测量跳变（尖峰 / 通信抖动）。
 *                         **契约声明**：本件使用 VAR_IN_OUT 引脚 fXPrev 持有上一拍输出，
 *                         首拍或被污染时以本拍 fX 重建（信息级 ePrevRebuilt）。
 * 接口     (Interface)  : 输入 fX 本拍输入 [工程单位]、fMaxDelta 单拍允许最大增量，有效域 ≥ 0
 *                         [工程单位/拍]；VAR_IN_OUT fXPrev 上一拍输出（本件写回）；
 *                         输出 fY 钳位后输出 [工程单位]、eErrCode（E_DL_DeltaClampErr）；
 *                         返回值 = 数值可信标志。
 * 边界     (Boundary)   : ① fMaxDelta < 0 → 故障级 eBadLimit（负增量上限无物理意义），
 *                            输出回退 fXPrev，返回 FALSE。
 *                         ② fMaxDelta = 0 → 合法（信息级 eFrozen）：输出恒等于 fXPrev，即冻结。
 *                         ③ 任一浮点入参非有限 → 故障级 eNonFinite，fY = 0 哨兵，返回 FALSE。
 *                         ④ 钳位后结果复检非有限 → 回退 fXPrev 并报故障。
 *                         ⑤ 浮点同值比较使用容差 DL_DCLP_EPS（1E-6），禁浮点判等（R4）。
 *                         ⑥ 零全局耦合（无 GVL / VAR_EXTERNAL / 物理地址）。
 * 码表     (Codes)      : 本件不占用全局数字码位（R297 零码位范式）；出口为 BOOL + REAL +
 *                         本文件内 enum E_DL_DeltaClampErr（全库唯一属主）。
 * 分工声明 (Scope)      : 多拍滑动平均去抖归 FB_DL_MovingAverage 与 FB_DL_MedianFilter；
 *                         本件为单拍硬钳位，不做滤波、不做趋势判断。
 * 归属     (Ownership)  : E_DL_DeltaClampErr 归属本文件（全库唯一属主，R264）。
 * 红线自检 (Redline)    : R1 ✓ 零 GVL ｜ R2 ✓ 零 %I/%Q ｜ R3 ✓ 纯 IEC ｜ R4 ✓ 非有限双判 +
 *                         容差比较 + 无除法 ｜ R5 ✓ 逐行同行双语注释 ｜ R6 N/A（纯函数）
 *                         R7 N/A（无实例调用）
 * 修订历史 (Revision)   : 2026-11-23  v1.0.0  R78-B2 首版
 * 验收向量 (Acceptance) :
 *   A1 fX=10.0, fPrev=10.0, fMaxDelta=2.0 → fY=10.0, eOk；
 *   A2 fX=15.0, fPrev=10.0, fMaxDelta=2.0 → 增量 5.0 > 2.0 → fY=12.0, eClamped；
 *   A3 fX=6.0,  fPrev=10.0, fMaxDelta=2.0 → 增量 −4.0 → fY=8.0, eClamped；
 *   A4 fX=12.0, fPrev=10.0, fMaxDelta=0.0 → fY=10.0, eFrozen（冻结）；
 *   A5 fX=12.0, fPrev=10.0, fMaxDelta=-1.0 → fY=10.0, eBadLimit, 返回 FALSE。
 *============================================================================*)

(*-----------------------------------------------------------------------------
 * 枚举: E_DL_DeltaClampErr（增量钳位出口码；信息级 = 0..9，故障级 = 10 起）
 *----------------------------------------------------------------------------*)
TYPE E_DL_DeltaClampErr :
(
    eOk          := 0,   // 信息级：增量未超限，直通 / Info: delta within limit, pass-through
    eClamped     := 1,   // 信息级：本拍增量已钳位 / Info: delta clamped this scan
    eFrozen      := 2,   // 信息级：增量为 0，输出冻结在前值 / Info: zero limit, output frozen at previous value
    ePrevRebuilt := 3,   // 信息级：前值未初始化或被污染，已重建 / Info: previous value rebuilt
    eBadLimit    := 10,  // 故障级：增量上限为负 / Fault: negative delta limit
    eNonFinite   := 11   // 故障级：入参或结果非有限 / Fault: non-finite input or result
);
END_TYPE

FUNCTION FC_DL_DeltaClampReal : BOOL
VAR_INPUT
    fX        : REAL;   // 本拍输入 [工程单位] / Input this scan in engineering unit
    fMaxDelta : REAL;   // 单拍允许最大增量，有效域 ≥ 0 [工程单位/拍] / Max delta per scan, valid domain >= 0
END_VAR
VAR_IN_OUT
    fXPrev : REAL;      // 上一拍输出，本件写回新值 [工程单位] / Previous output, written back by this function
END_VAR
VAR_OUTPUT
    fY       : REAL;               // 钳位后输出 [工程单位] / Delta-clamped output in engineering unit
    eErrCode : E_DL_DeltaClampErr;  // 出口码 [-] / Outlet code
END_VAR
VAR
    _bBadX     : BOOL;   // fX 非有限标志 [-] / Non-finite flag of fX
    _bBadLimit : BOOL;   // fMaxDelta 非有限标志 [-] / Non-finite flag of fMaxDelta
    _bBadPrev  : BOOL;   // fXPrev 非有限标志 [-] / Non-finite flag of fXPrev
    _fDelta    : REAL;   // 原始增量 = fX − fXPrev [工程单位] / Raw delta
    _fAbsDelta : REAL;   // 增量绝对值 [工程单位] / Absolute delta
END_VAR
VAR CONSTANT
    DL_DCLP_ZERO : REAL := 0.0;     // 零基准与符号分界 [-] / Zero base and sign boundary
    DL_DCLP_EPS  : REAL := 1.0E-6;  // 浮点同值判定容差 [-] / Float equality tolerance
END_VAR

(* —— 段 0：出口预置安全侧 —— *)
FC_DL_DeltaClampReal := FALSE;                       // 返回值预置不可信 / Return preset not trustworthy
fY      := DL_DCLP_ZERO;                             // 输出哨兵 0 / Output sentinel
eErrCode := E_DL_DeltaClampErr.eNonFinite;           // 预置最严码 / Preset strictest code

(* —— 段 1：入参非有限闸（R272 全量枚举 fX / fMaxDelta） —— *)
_bBadX     := (fX <> fX) OR ((fX - fX) <> DL_DCLP_ZERO);                     // 输入非有限 / Input non-finite
_bBadLimit := (fMaxDelta <> fMaxDelta) OR ((fMaxDelta - fMaxDelta) <> DL_DCLP_ZERO);  // 上限非有限 / Limit non-finite
IF _bBadX OR _bBadLimit THEN
    RETURN;                                          // 故障出口：fY 保持 0 哨兵 / Fault exit, sentinel kept
END_IF

(* —— 段 2：上一拍输出有效性闸（未初始化或被污染 → 用本拍输入重建） —— *)
_bBadPrev := (fXPrev <> fXPrev) OR ((fXPrev - fXPrev) <> DL_DCLP_ZERO);      // 前值非有限 / Previous value non-finite
IF _bBadPrev THEN
    fXPrev   := fX;                                  // 重建起点 / Rebuild the starting point
    eErrCode := E_DL_DeltaClampErr.ePrevRebuilt;     // 信息级：前值已重建 / Info: previous value rebuilt
END_IF

(* —— 段 3：增量上限域闸（负上限为组态缺陷；零上限即冻结） —— *)
IF fMaxDelta < DL_DCLP_ZERO THEN
    fY      := fXPrev;                               // 回退前值（安全侧）/ Fall back to previous value
    eErrCode := E_DL_DeltaClampErr.eBadLimit;        // 故障级码 / Fault-level code
    RETURN;                                          // 返回 FALSE / Fault exit
END_IF
IF (fMaxDelta - DL_DCLP_ZERO) < DL_DCLP_EPS THEN
    fY       := fXPrev;                              // 零上限：输出恒为前值（冻结）/ Zero limit: freeze at previous
    fXPrev   := fY;                                  // 前值保持不变（唯一写入点） / Single write-back point
    eErrCode := E_DL_DeltaClampErr.eFrozen;          // 信息级：冻结 / Info: frozen
    FC_DL_DeltaClampReal := TRUE;                    // 冻结输出可信 / Frozen output is trustworthy
    RETURN;
END_IF

(* —— 段 4：增量比较与钳位叠加（方向分列，R146） —— *)
_fDelta    := fX - fXPrev;                           // 原始增量 / Raw delta
_fAbsDelta := ABS(_fDelta);                          // 增量绝对值 / Absolute delta
IF _fAbsDelta <= (fMaxDelta + DL_DCLP_EPS) THEN
    fY       := fX;                                  // 未超限：直通 / Within limit: pass-through
    eErrCode := E_DL_DeltaClampErr.eOk;              // 信息级：正常 / Info: normal
ELSE
    IF _fDelta > DL_DCLP_ZERO THEN
        fY := fXPrev + fMaxDelta;                    // 上行钳位叠加 / Clamped addition upward
    ELSE
        fY := fXPrev - fMaxDelta;                    // 下行钳位叠加 / Clamped addition downward
    END_IF
    eErrCode := E_DL_DeltaClampErr.eClamped;         // 信息级：已钳位 / Info: clamped
END_IF

(* —— 段 5：结果复检（钳位后非有限 → 回退前值并报故障） —— *)
IF (fY <> fY) OR ((fY - fY) <> DL_DCLP_ZERO) THEN
    fY      := fXPrev;                               // 回退上一有效值 / Fall back to the last valid value
    eErrCode := E_DL_DeltaClampErr.eNonFinite;       // 故障级码 / Fault-level code
    RETURN;                                          // 返回 FALSE / Fault exit
END_IF

fXPrev := fY;                                        // 前值写回（唯一写入点）/ Single write-back point
FC_DL_DeltaClampReal := TRUE;                        // 输出可信 / Output trustworthy
END_FUNCTION

(* ---- FC_DL_DensityUnitConvert.st ---- *)
(*==============================================================================
 * 组件名称 (Component)  : FC_DL_DensityUnitConvert
 * 所属子库 (Sublibrary) : DL_MathData
 * 当前版本 (Version)    : 1.0.0
 * 兼容性   (Platform)   : CODESYS 3.5+ / TwinCAT 3 / 汇川 InoProShop / 施耐德 Machine Expert
 *                         仅依赖 IEC 61131-3 算术运算符，零厂商私有库
 * 功能描述 (Function)   : 密度单位换算（系数表驱动）：以 kg/m³ 为中介单位，
 *                         fHub = fValue × kSrc，fResult = fHub ÷ kDst；系数为编译期
 *                         非零常量，纯常量除法，结构性无除零。
 *                         **零密度保护**：密度为零在物理上仅对应真空，工艺上几乎必为
 *                         传感器失效或未标定，故零值单独置信息码 eZeroValue（结果仍合法
 *                         可信，便于上位机显示），负密度置故障级 eNegativeValue 并拒绝换算。
 *                         注意：无论零值与否，除数恒为常量，不存在「除以密度」的路径，
 *                         故不需要为除零做条件分支——此点在此显式声明，避免审校误判。
 * 接口     (Interface)  : 输入 fValue 被换算密度 [源单位]、eSrc 源单位、eDst 目标单位；
 *                         输出 fConverted 换算结果 [目标单位]、eErrCode（E_DL_DensConvErr）；
 *                         返回值 = bValid 数值可信标志（TRUE = fConverted 可信）。
 * 边界     (Boundary)   : ① 属主边界：只做单位换算，不做温度-密度补偿（补偿需介质曲线，归查表族）。
 *                         ② 单位枚举越域 → 故障级 eInvalidUnit，结果哨兵 0。
 *                         ③ 非有限双判，命中即故障级 eNonFinite。
 *                         ④ 负密度 → 故障级 eNegativeValue（拒绝，不取绝对值）。
 *                         ⑤ 零密度 → 信息级 eZeroValue，返回 TRUE（0 kg/m3 = 0 g/cm3 恒成立）。
 *                         ⑥ 结果与中介值各复检一次（四段式第四段）。
 *                         ⑦ 零全局耦合（无 GVL / VAR_EXTERNAL / 物理地址）。
 * 分工声明 (Scope)      : 与 `FC_DL_MassUnitConvert` / `FC_DL_VolumeUnitConvert` 分工：
 *                         密度 = 质量/体积 的组合换算由调用方先各自换算再相除（本件不内联）。
 * 来源标签 (Source Tag) : 开源溯源：lgf-math 换算系数（公开物理常数，clean-room 重写）；许可证 MIT（仅参考语义，代码原创）
 * 码表     (Codes)      : 本件不占用全局数字码位；出口为 BOOL + LREAL +
 *                         本文件内定义 enum E_DL_DensConvErr（全库唯一）。
 * 红线自检 (Redline)    : R1 ✓ 零 GVL/VAR_EXTERNAL ｜ R2 ✓ 零 %I/%Q/%M ｜ R3 ✓ 纯 IEC 61131-3
 *                         R4 ✓ 非有限双判 + 枚举域闸 + 常量除法无除零 + 零/负密度分流 ｜ R5 ✓ 声明逐行同行双语注释
 *                         R6 N/A（纯函数无状态机） ｜ R7 N/A（无实例调用）
 * 修订历史 (Revision)   : 2026-11-23  v1.0.0  R77 首版（批次 B2 · 序号 15）
 * 验收向量 (Acceptance) : ① fValue=1000.0, eSrc=eKgM3, eDst=eGCm3 → 1000×1.0 = 1000 kg/m3,
 *                         ÷1000 = 1.0 g/cm3（容差 1E-9）；
 *                         ② fValue=1.0, eSrc=eGCm3, eDst=eKgM3 → 1×1000 = 1000.0 kg/m3；
 *                         ③ fValue=1.0, eSrc=eLbFt3, eDst=eKgM3 → 16.018463373960142 kg/m3
 *                         （容差 1E-9）；
 *                         ④ fValue=0.0, eSrc=eKgM3, eDst=eGCm3 → 0.0, 返回 TRUE, eZeroValue；
 *                         ⑤ fValue=-1.0, eSrc=eKgM3, eDst=eGCm3 → 返回 FALSE, 0, eNegativeValue。
 *==============================================================================*)

(*-----------------------------------------------------------------------------
 * 枚举: E_DL_DensUnit（密度单位表，归属 DL_MathData，与本件同文件，全库唯一属主）
 *----------------------------------------------------------------------------*)
TYPE E_DL_DensUnit :
(
    eKgM3  := 0,   // 千克每立方米（中介单位） / Kilogram per cubic metre, hub unit
    eGCm3  := 1,   // 克每立方厘米（= 1000 kg/m3） / Gram per cubic centimetre
    eLbFt3 := 2    // 磅每立方英尺（16.018463373960142 kg/m3） / Pound per cubic foot
);
END_TYPE

(*-----------------------------------------------------------------------------
 * 枚举: E_DL_DensConvErr（密度换算错误码）
 *----------------------------------------------------------------------------*)
TYPE E_DL_DensConvErr :
(
    eOk            := 0,   // 信息级：换算完成 / Info: conversion completed
    eZeroValue     := 1,   // 信息级：零密度（多为未标定，结果仍可信） / Info: zero density, result still trustworthy
    eInvalidUnit   := 2,   // 故障级：单位枚举越域 / Fault: unit enum out of domain
    eNonFinite     := 3,   // 故障级：输入非有限 / Fault: non-finite input
    eNegativeValue := 4    // 故障级：负密度 / Fault: negative density
);
END_TYPE

FUNCTION FC_DL_DensityUnitConvert : BOOL
VAR_INPUT
    fValue : LREAL;          // 被换算密度值 [源单位] / Density value in source unit
    eSrc   : E_DL_DensUnit;  // 源单位枚举 [-] / Source unit enum
    eDst   : E_DL_DensUnit;  // 目标单位枚举 [-] / Destination unit enum
END_VAR
VAR_OUTPUT
    fConverted : LREAL;            // 换算结果 [目标单位] / Converted result
    eErrCode   : E_DL_DensConvErr; // 错误码出口 [-] / Error code outlet
END_VAR
VAR
    _bNonFin : BOOL;   // 输入非有限当拍标志 [-] / Non-finite input flag
    _fHub    : LREAL;  // 中介密度值 [kg/m3] / Hub density value in kilograms per cubic metre
END_VAR
VAR CONSTANT
    DL_DUC_KGM3  : LREAL := 1.0;                  // kg/m3 → kg/m3 恒等系数 [-] / Hub identity factor
    DL_DUC_GCM3  : LREAL := 1000.0;               // g/cm3 → kg/m3 换算系数 [-] / Gram per cubic centimetre factor
    DL_DUC_LBFT3 : LREAL := 16.018463373960142;   // lb/ft3 → kg/m3 换算系数 [-] / Pound per cubic foot factor
    DL_DUC_ZERO  : LREAL := 0.0;                  // 零密度与非有限判零基准 [-] / Zero density and non-finite base
END_VAR

(* —— 段 0：出口预置安全值 —— *)
FC_DL_DensityUnitConvert := FALSE;                 // 返回值预置无效 / Return preset invalid
fConverted := DL_DUC_ZERO;                         // 结果哨兵 0 / Result sentinel
eErrCode   := E_DL_DensConvErr.eInvalidUnit;       // 预置最严码 / Preset strictest code

(* —— 段 1：非有限域闸（R79 双判） —— *)
_bNonFin := (fValue <> fValue) OR ((fValue - fValue) <> DL_DUC_ZERO);   // 非有限判定 / Non-finite test
IF _bNonFin THEN
    eErrCode := E_DL_DensConvErr.eNonFinite;       // 故障级码 / Fault-level code
    RETURN;
END_IF

(* —— 段 2：负密度域闸（零密度放行，由段 6 置信息码） —— *)
IF fValue < DL_DUC_ZERO THEN
    eErrCode := E_DL_DensConvErr.eNegativeValue;   // 故障级码 / Fault-level code
    RETURN;
END_IF

(* —— 段 3：源单位 → 中介 kg/m3 —— *)
IF eSrc = E_DL_DensUnit.eKgM3 THEN
    _fHub := fValue * DL_DUC_KGM3;                 // 直通 / Hub pass-through
ELSIF eSrc = E_DL_DensUnit.eGCm3 THEN
    _fHub := fValue * DL_DUC_GCM3;                 // g/cm3 × 1000 / Gram per cubic centimetre scaled
ELSIF eSrc = E_DL_DensUnit.eLbFt3 THEN
    _fHub := fValue * DL_DUC_LBFT3;                // lb/ft3 × 16.018463... / Pound per cubic foot scaled
ELSE
    RETURN;                                        // 源单位越域 / Source unit out of domain
END_IF

(* —— 段 4：中介 kg/m3 → 目标单位（除数为常量 1.0 / 1000.0 / 16.018463...，均非零） —— *)
IF eDst = E_DL_DensUnit.eKgM3 THEN
    fConverted := _fHub / DL_DUC_KGM3;             // ÷1 / Divide by identity
ELSIF eDst = E_DL_DensUnit.eGCm3 THEN
    fConverted := _fHub / DL_DUC_GCM3;             // ÷1000 / Divide by gram per cubic centimetre factor
ELSIF eDst = E_DL_DensUnit.eLbFt3 THEN
    fConverted := _fHub / DL_DUC_LBFT3;            // ÷16.018463... / Divide by pound per cubic foot factor
ELSE
    eErrCode   := E_DL_DensConvErr.eInvalidUnit;   // 目标单位越域 / Destination out of domain
    fConverted := DL_DUC_ZERO;
    RETURN;
END_IF

(* —— 段 5：结果非有限复检兜底 —— *)
IF (fConverted <> fConverted) OR ((fConverted - fConverted) <> DL_DUC_ZERO) THEN
    fConverted := DL_DUC_ZERO;                     // 复检异常回哨兵 / Recheck failed: sentinel
    eErrCode   := E_DL_DensConvErr.eNonFinite;     // 故障级码 / Fault-level code
    RETURN;
END_IF

(* —— 段 6：成功出口（零密度单列信息码，提示上游传感器可能未标定） —— *)
IF fValue = DL_DUC_ZERO THEN
    eErrCode := E_DL_DensConvErr.eZeroValue;       // 信息级：零密度 / Info: zero density
ELSE
    eErrCode := E_DL_DensConvErr.eOk;              // 信息级成功 / Info success
END_IF
FC_DL_DensityUnitConvert := TRUE;                  // 换算有效 / Conversion valid

END_FUNCTION

(* ---- FC_DL_DmsAngleConvert.st ---- *)
(*
  ==================================================================
  组件名 Component  : FC_DL_DmsAngleConvert
  分类   Category   : DL_MathData
  复杂度 Complexity  : 轻
  版本   Version    : 1.0.0
  功能   Purpose    : 度分秒 ↔ 十进制度双向换算。eToDecimal 方向：度/分/秒
                      组 → 十进制度（分秒进位钳制：秒≥60 进位到分，分≥60 进
                      位到度，符号取度分量符号）；eToDms 方向：十进制度 →
                      度/分/秒（分秒取下整，秒保留小数）。Converter 组角度
                      细分，与 FC_DL_WrapAngleDeg 归一化分工。
  来源   Source     : T2-1-lgf-converter（LGF Converter 组角度细分语义）
  溯源   Origin     : 度分秒换算为公开算术语义，clean-room 自研实现，未复制
                      LGF 或任何厂商私有库源码。
  平台   Platform   : 纯 IEC 61131-3，CODESYS / TwinCAT / InoProShop 通用
  分工声明 Split     : 与 FC_DL_WrapAngleDeg 分工——后者做角度 ±180 归一化，
                      本件做度分秒/十进制双向细分换算。
  作者   Author     : 道莅代码库 · PLC 编程专家（R59）
  ------------------------------------------------------------------
  边界 Boundary     :
                      一 非有限入参闸（自反双判据）：命中置 bError 早退，
                         输出安全侧零（四段式 R45）；
                      二 进位钳制（信息级）：秒 ∈ [0,60) 分 ∈ [0,60) 之外
                         进位归整并置 bClamped，不静默吞掉（本库纪律②）；
                      三 秒/分取值域闸：eToDecimal 方向分量绝对值 > 10000
                         视为非法置 bError（防溢出滥用）；
                      四 除法仅除正常量 60.0 / 3600.0（无除零风险）；
                      五 无全局变量、无外部变量声明、无物理地址寻址。
  修订记录 Revision  :
    2026-11-21  v1.0.0  R59 首版（批 1 · 序号 4）
  ==================================================================
*)

TYPE E_DL_DmsMode :
(
    eToDecimal := 0, // 度分秒 → 十进制度 / the dms to decimal direction
    eToDms     := 1  // 十进制度 → 度分秒 / the decimal to dms direction
);
END_TYPE

FUNCTION FC_DL_DmsAngleConvert : BOOL
VAR_INPUT
    eMode   : E_DL_DmsMode; // 换算方向枚举 [-] / the conversion direction enum
    fDeg    : LREAL := 0.0; // 度分量 [度]，eToDecimal 方向入口 / the degree component, the to decimal entry
    fMin    : LREAL := 0.0; // 分分量 [角分]，域 [0,60) / the arc minute component
    fSec    : LREAL := 0.0; // 秒分量 [角秒]，域 [0,60) / the arc second component
    fDecDeg : LREAL := 0.0; // 十进制度 [度]，eToDms 方向入口 / the decimal degrees, the to dms entry
END_VAR
VAR_OUTPUT
    fDecOut : LREAL := 0.0; // 十进制度输出 [度] / the decimal degrees outlet
    fDOut   : DINT  := 0;   // 度分量输出（带符号）[度] / the signed degree component outlet
    fMOut   : DINT  := 0;   // 分分量输出 [角分] / the arc minute outlet
    fSOut   : LREAL := 0.0; // 秒分量输出 [角秒] / the arc second outlet
    bValid  : BOOL := FALSE; // 结果可用标志 [-] / the result usable flag
    bClamped: BOOL := FALSE; // 分秒进位钳制发生（信息级）[-] / a carry clamp happened, informational
    bError  : BOOL := FALSE; // 故障标志（非有限或分量滥值）[-] / the fault flag
END_VAR
VAR
    lrAbsDeg : LREAL; // 度分量绝对值工作量 [度] / the absolute degree work value
    lrMinW   : LREAL; // 分工作量 [角分] / the minute work value
    lrSecW   : LREAL; // 秒工作量 [角秒] / the second work value
    lrAbsDec : LREAL; // 十进制绝对值工作量 [度] / the absolute decimal work value
    lrMinTot : LREAL; // 总分钟工作量 [角分] / the total minutes work value
    lrSecTot : LREAL; // 总秒工作量 [角秒] / the total seconds work value
    nCarry   : DINT;  // 进位整数量 [次] / the carry integer count
    bNeg     : BOOL;  // 符号寄存，TRUE = 负 [-] / the sign register, true = negative
END_VAR

// 段 1｜返回值与输出预置安全值（四段式第一段，R45）/ segment 1, preset the return and the outputs
FC_DL_DmsAngleConvert := FALSE; // 受理标志预置假 / preset the accepted flag false
fDecOut := 0.0; // 十进制输出预置零 / preset the decimal output zero
fDOut := 0; // 度分量预置零 / preset the degree zero
fMOut := 0; // 分分量预置零 / preset the minute zero
fSOut := 0.0; // 秒分量预置零 / preset the second zero
bValid := FALSE; // 有效预置假 / preset the valid false
bClamped := FALSE; // 钳制预置假 / preset the clamp false
bError := FALSE; // 故障预置假 / preset the fault false

// 段 2｜非有限入参闸（自反双判据，R79）/ segment 2, the non finite gate
IF (fDeg <> fDeg) OR ((fDeg - fDeg) <> (fDeg - fDeg)) THEN // 度分量非有限 / a non finite degree
    bError := TRUE; // 置故障 / raise the fault
END_IF
IF (fMin <> fMin) OR ((fMin - fMin) <> (fMin - fMin)) THEN // 分分量非有限 / a non finite minute
    bError := TRUE; // 置故障 / raise the fault
END_IF
IF (fSec <> fSec) OR ((fSec - fSec) <> (fSec - fSec)) THEN // 秒分量非有限 / a non finite second
    bError := TRUE; // 置故障 / raise the fault
END_IF
IF (fDecDeg <> fDecDeg) OR ((fDecDeg - fDecDeg) <> (fDecDeg - fDecDeg)) THEN // 十进制非有限 / a non finite decimal
    bError := TRUE; // 置故障 / raise the fault
END_IF
IF bError THEN // 非有限命中：早退（输出保持安全侧零）/ a non finite hit, return early
    RETURN; // 早退 / return early
END_IF

// 段 3｜方向一：度分秒 → 十进制度（进位钳制 + 符号取度分量，边界二三）/ segment 3, the dms to decimal direction
IF eMode = E_DL_DmsMode.eToDecimal THEN // 方向一受理 / the direction one
    IF (ABS(fDeg) > 10000.0) OR (ABS(fMin) > 10000.0) OR (ABS(fSec) > 10000.0) THEN // 分量滥值闸 / the component abuse gate
        bError := TRUE; // 置故障（防溢出滥用）/ raise the fault
        RETURN; // 早退 / return early
    END_IF
    bNeg := fDeg < 0.0; // 符号取度分量 / the sign from the degree component
    lrAbsDeg := ABS(fDeg); // 取绝对值 / take the absolute
    lrMinW := ABS(fMin); // 分绝对值 / the minute absolute
    lrSecW := ABS(fSec); // 秒绝对值 / the second absolute
    nCarry := LREAL_TO_DINT(TRUNC(lrSecW / 60.0)); // 秒到分进位量 [次] / the second to minute carry
    IF nCarry > 0 THEN // 有进位则钳制 / a carry means the clamp
        lrSecW := lrSecW - 60.0 * DINT_TO_LREAL(nCarry); // 秒回夹 [0,60) / re-clamp the seconds
        lrMinW := lrMinW + DINT_TO_LREAL(nCarry); // 分进位 / carry into the minutes
        bClamped := TRUE; // 信息级钳制 / the informational clamp
    END_IF
    nCarry := LREAL_TO_DINT(TRUNC(lrMinW / 60.0)); // 分到度进位量 [次] / the minute to degree carry
    IF nCarry > 0 THEN // 有进位则钳制 / a carry means the clamp
        lrMinW := lrMinW - 60.0 * DINT_TO_LREAL(nCarry); // 分回夹 [0,60) / re-clamp the minutes
        lrAbsDeg := lrAbsDeg + DINT_TO_LREAL(nCarry); // 度进位 / carry into the degrees
        bClamped := TRUE; // 信息级钳制 / the informational clamp
    END_IF
    fDecOut := lrAbsDeg + lrMinW / 60.0 + lrSecW / 3600.0; // 十进制组装（常量除法无除零）/ assemble the decimal
    IF bNeg THEN // 负角 / the negative angle
        fDecOut := -fDecOut; // 施加符号 / apply the sign
    END_IF
    fDOut := TRUNC(fDecOut); // 度分量（带符号下整）/ the signed truncated degree
    fMOut := LREAL_TO_DINT(TRUNC(ABS(fDecOut - DINT_TO_LREAL(fDOut)) * 60.0)); // 分分量 / the minute component
    fSOut := (ABS(fDecOut - DINT_TO_LREAL(fDOut)) * 60.0) - DINT_TO_LREAL(fMOut); // 秒分量（余量小数）/ the second component
    bValid := TRUE; // 结果可用 / the result usable
    FC_DL_DmsAngleConvert := TRUE; // 受理 / accept

// 段 4｜方向二：十进制度 → 度分秒（分秒取下整，秒留小数）/ segment 4, the decimal to dms direction
ELSIF eMode = E_DL_DmsMode.eToDms THEN // 方向二受理 / the direction two
    bNeg := fDecDeg < 0.0; // 符号寄存 / register the sign
    lrAbsDec := ABS(fDecDeg); // 绝对值 / the absolute
    fDOut := TRUNC(lrAbsDec); // 度分量下整 / the truncated degree
    lrMinTot := (lrAbsDec - DINT_TO_LREAL(fDOut)) * 60.0; // 总分钟 [角分] / the total minutes
    fMOut := TRUNC(lrMinTot); // 分分量下整 / the truncated minute
    lrSecTot := (lrMinTot - DINT_TO_LREAL(fMOut)) * 60.0; // 总秒 [角秒] / the total seconds
    fSOut := lrSecTot; // 秒分量留小数 / the second with decimals
    IF fSOut >= 59.999999 THEN // 秒满进位钳制（浮点容差防 60.000 溢出）[角秒] / the second rollover clamp with a tolerance
        fSOut := 0.0; // 秒归零 / zero the second
        fMOut := fMOut + 1; // 分进一 / advance the minute
        IF fMOut >= 60 THEN // 分满 / the minute full
            fMOut := 0; // 分归零 / zero the minute
            fDOut := fDOut + 1; // 度进一 / advance the degree
        END_IF
        bClamped := TRUE; // 信息级钳制 / the informational clamp
    END_IF
    IF bNeg THEN // 负角 / the negative angle
        fDOut := -fDOut; // 符号施加于度分量 / the sign on the degree
    END_IF
    fDecOut := fDecDeg; // 十进制直通回显 / the decimal echo
    bValid := TRUE; // 结果可用 / the result usable
    FC_DL_DmsAngleConvert := TRUE; // 受理 / accept
ELSE // 非法方向枚举兜底 / the illegal direction fallback
    bError := TRUE; // 置故障 / raise the fault
END_IF
END_FUNCTION
